Universal Robots URScript: FaiChun_9 Jan_3.script

def Machining1():
  # Default parameters:
  global speed_ms = 0.03
  global speed_rads = 0.75
  global accel_mss = 3
  global accel_radss = 1.2
  global blend_radius_m = 0.0003

  # Add subprograms here
  # Start of main program
  # Program generated by RoboDK v5.6.8 for UR10e on 09/01/2025 16:15:55
  # Using nominal kinematics.
  blend_radius_m = 0.0003
  speed_ms = 0.03
  # set_reference(p[0.335000, -0.060000, 0.000000, 0.000000, 0.000000, 0.000000])
  set_tcp(p[0.000000, 0.000000, 0.252000, 0.000000, 0.000000, 0.000000])
  # Show Tool
  movej([0.602689, -1.119966, -2.613047, -0.979376, 1.570796, 2.173486],accel_radss,speed_rads,0,blend_radius_m)
  movel([0.602689, -1.179994, -2.651340, -0.881054, 1.570796, 2.173486],accel_mss,speed_ms,0,blend_radius_m)
  #SetTool1
  #M_RunCode6
  #SetRPM60000
  speed_ms = 0.03
  #M_RunCode3
  movel([0.602689, -1.207513, -2.665873, -0.839003, 1.570796, 2.173486],accel_mss,speed_ms,0,blend_radius_m)
  speed_ms = 0.003
  movel([0.602689, -1.214750, -2.669441, -0.828198, 1.570796, 2.173486],accel_mss,speed_ms,0,blend_radius_m)
  speed_ms = 0.007
  movel([0.623056, -1.305978, -2.619553, -0.786857, 1.570796, 2.193852],accel_mss,speed_ms,0,blend_radius_m)
  movel([0.614868, -1.310439, -2.616847, -0.785103, 1.570796, 2.185664],accel_mss,speed_ms,0,blend_radius_m)
  movel([0.615927, -1.315223, -2.613916, -0.783250, 1.570796, 2.186723],accel_mss,speed_ms,0,blend_radius_m)
  movel([0.618034, -1.314081, -2.614619, -0.783689, 1.570796, 2.188830],accel_mss,speed_ms,0,blend_radius_m)
  movel([0.617346, -1.310924, -2.616551, -0.784913, 1.570796, 2.188143],accel_mss,speed_ms,0,blend_radius_m)
  movel([0.623401, -1.307643, -2.618547, -0.786200, 1.570796, 2.194198],accel_mss,speed_ms,0,blend_radius_m)
  movel([0.623560, -1.308410, -2.618081, -0.785898, 1.570796, 2.194357],accel_mss,speed_ms,0,blend_radius_m)
  movel([0.624387, -1.312349, -2.615681, -0.784359, 1.570796, 2.195184],accel_mss,speed_ms,0,blend_radius_m)
  movel([0.620317, -1.314540, -2.614336, -0.783512, 1.570796, 2.191113],accel_mss,speed_ms,0,blend_radius_m)
  movel([0.620668, -1.316175, -2.613329, -0.782885, 1.570796, 2.191464],accel_mss,speed_ms,0,blend_radius_m)
  movel([0.624731, -1.313996, -2.614671, -0.783722, 1.570796, 2.195527],accel_mss,speed_ms,0,blend_radius_m)
  movel([0.625701, -1.318667, -2.611788, -0.781935, 1.570796, 2.196498],accel_mss,speed_ms,0,blend_radius_m)
  movel([0.621661, -1.320822, -2.610447, -0.781120, 1.570796, 2.192457],accel_mss,speed_ms,0,blend_radius_m)
  movel([0.622322, -1.323943, -2.608496, -0.779950, 1.570796, 2.193118],accel_mss,speed_ms,0,blend_radius_m)
  movel([0.616386, -1.327108, -2.606503, -0.778778, 1.570796, 2.187182],accel_mss,speed_ms,0,blend_radius_m)
  movel([0.615701, -1.324013, -2.608452, -0.779924, 1.570796, 2.186497],accel_mss,speed_ms,0,blend_radius_m)
  movel([0.613619, -1.325132, -2.607748, -0.779508, 1.570796, 2.184416],accel_mss,speed_ms,0,blend_radius_m)
  movel([0.614310, -1.328222, -2.605799, -0.778369, 1.570796, 2.185106],accel_mss,speed_ms,0,blend_radius_m)
  movel([0.609368, -1.330876, -2.604114, -0.777400, 1.570796, 2.180164],accel_mss,speed_ms,0,blend_radius_m)
  movel([0.608412, -1.331392, -2.603784, -0.777212, 1.570796, 2.179209],accel_mss,speed_ms,0,blend_radius_m)
  movel([0.607352, -1.326855, -2.606663, -0.778871, 1.570796, 2.178148],accel_mss,speed_ms,0,blend_radius_m)
  movel([0.611354, -1.324685, -2.608029, -0.779674, 1.570796, 2.182150],accel_mss,speed_ms,0,blend_radius_m)
  movel([0.610987, -1.323080, -2.609036, -0.780272, 1.570796, 2.181784],accel_mss,speed_ms,0,blend_radius_m)
  movel([0.604903, -1.326389, -2.606957, -0.779043, 1.570796, 2.175699],accel_mss,speed_ms,0,blend_radius_m)
  movel([0.606349, -1.332504, -2.603075, -0.776810, 1.570796, 2.177146],accel_mss,speed_ms,0,blend_radius_m)
  movel([0.503740, -1.390840, -2.563439, -0.758110, 1.570796, 2.074536],accel_mss,speed_ms,0,blend_radius_m)
  movel([0.410742, -1.448915, -2.519079, -0.744396, 1.570796, 1.981539],accel_mss,speed_ms,0,blend_radius_m)
  movel([0.408155, -1.444408, -2.522703, -0.745278, 1.570796, 1.978951],accel_mss,speed_ms,0,blend_radius_m)
  movel([0.403196, -1.447676, -2.520078, -0.744635, 1.570796, 1.973993],accel_mss,speed_ms,0,blend_radius_m)
  movel([0.403874, -1.448837, -2.519141, -0.744410, 1.570796, 1.974671],accel_mss,speed_ms,0,blend_radius_m)
  movel([0.407131, -1.446693, -2.520869, -0.744827, 1.570796, 1.977928],accel_mss,speed_ms,0,blend_radius_m)
  movel([0.409046, -1.450019, -2.518186, -0.744184, 1.570796, 1.979842],accel_mss,speed_ms,0,blend_radius_m)
  movel([0.408262, -1.450531, -2.517771, -0.744086, 1.570796, 1.979059],accel_mss,speed_ms,0,blend_radius_m)
  movel([0.404240, -1.453169, -2.515629, -0.743591, 1.570796, 1.975036],accel_mss,speed_ms,0,blend_radius_m)
  movel([0.402940, -1.450940, -2.517440, -0.744009, 1.570796, 1.973737],accel_mss,speed_ms,0,blend_radius_m)
  movel([0.401260, -1.452049, -2.516540, -0.743800, 1.570796, 1.972056],accel_mss,speed_ms,0,blend_radius_m)
  movel([0.402562, -1.454272, -2.514730, -0.743387, 1.570796, 1.973359],accel_mss,speed_ms,0,blend_radius_m)
  movel([0.397796, -1.457416, -2.512158, -0.742815, 1.570796, 1.968593],accel_mss,speed_ms,0,blend_radius_m)
  movel([0.396480, -1.455213, -2.513962, -0.743214, 1.570796, 1.967277],accel_mss,speed_ms,0,blend_radius_m)
  movel([0.393271, -1.457346, -2.512215, -0.742828, 1.570796, 1.964067],accel_mss,speed_ms,0,blend_radius_m)
  movel([0.391300, -1.454096, -2.514874, -0.743419, 1.570796, 1.962097],accel_mss,speed_ms,0,blend_radius_m)
  movel([0.394521, -1.451944, -2.516626, -0.743820, 1.570796, 1.965317],accel_mss,speed_ms,0,blend_radius_m)
  movel([0.393830, -1.450797, -2.517556, -0.744036, 1.570796, 1.964626],accel_mss,speed_ms,0,blend_radius_m)
  movel([0.390606, -1.452954, -2.515804, -0.743631, 1.570796, 1.961403],accel_mss,speed_ms,0,blend_radius_m)
  movel([0.388934, -1.450227, -2.518017, -0.744144, 1.570796, 1.959730],accel_mss,speed_ms,0,blend_radius_m)
  movel([0.388611, -1.449697, -2.518446, -0.744245, 1.570796, 1.959407],accel_mss,speed_ms,0,blend_radius_m)
  movel([0.393406, -1.446476, -2.521044, -0.744869, 1.570796, 1.964202],accel_mss,speed_ms,0,blend_radius_m)
  movel([0.394744, -1.448694, -2.519257, -0.744438, 1.570796, 1.965540],accel_mss,speed_ms,0,blend_radius_m)
  movel([0.396427, -1.447570, -2.520164, -0.744656, 1.570796, 1.967224],accel_mss,speed_ms,0,blend_radius_m)
  movel([0.394398, -1.444188, -2.522879, -0.745322, 1.570796, 1.965194],accel_mss,speed_ms,0,blend_radius_m)
  movel([0.387908, -1.448555, -2.519369, -0.744465, 1.570796, 1.958704],accel_mss,speed_ms,0,blend_radius_m)
  movel([0.387580, -1.448026, -2.519796, -0.744567, 1.570796, 1.958376],accel_mss,speed_ms,0,blend_radius_m)
  movel([0.348021, -1.388149, -2.565374, -0.758866, 1.570796, 1.918817],accel_mss,speed_ms,0,blend_radius_m)
  movel([0.300929, -1.326689, -2.606767, -0.778932, 1.570796, 1.871725],accel_mss,speed_ms,0,blend_radius_m)
  movel([0.308156, -1.320668, -2.610543, -0.781178, 1.570796, 1.878952],accel_mss,speed_ms,0,blend_radius_m)
  movel([0.305290, -1.317157, -2.612722, -0.782509, 1.570796, 1.876086],accel_mss,speed_ms,0,blend_radius_m)
  movel([0.303402, -1.318735, -2.611745, -0.781909, 1.570796, 1.874198],accel_mss,speed_ms,0,blend_radius_m)
  movel([0.305295, -1.321037, -2.610313, -0.781039, 1.570796, 1.876092],accel_mss,speed_ms,0,blend_radius_m)
  movel([0.299947, -1.325499, -2.607518, -0.779372, 1.570796, 1.870743],accel_mss,speed_ms,0,blend_radius_m)
  movel([0.299492, -1.324951, -2.607863, -0.779576, 1.570796, 1.870288],accel_mss,speed_ms,0,blend_radius_m)
  movel([0.297126, -1.322128, -2.609632, -0.780629, 1.570796, 1.867922],accel_mss,speed_ms,0,blend_radius_m)
  movel([0.300740, -1.319092, -2.611523, -0.781773, 1.570796, 1.871536],accel_mss,speed_ms,0,blend_radius_m)
  movel([0.299747, -1.317902, -2.612261, -0.782225, 1.570796, 1.870544],accel_mss,speed_ms,0,blend_radius_m)
  movel([0.296130, -1.320947, -2.610369, -0.781072, 1.570796, 1.866927],accel_mss,speed_ms,0,blend_radius_m)
  movel([0.293273, -1.317580, -2.612461, -0.782348, 1.570796, 1.864069],accel_mss,speed_ms,0,blend_radius_m)
  movel([0.296899, -1.314508, -2.614356, -0.783525, 1.570796, 1.867695],accel_mss,speed_ms,0,blend_radius_m)
  movel([0.294961, -1.312214, -2.615763, -0.784412, 1.570796, 1.865757],accel_mss,speed_ms,0,blend_radius_m)
  movel([0.300378, -1.307616, -2.618562, -0.786210, 1.570796, 1.871174],accel_mss,speed_ms,0,blend_radius_m)
  movel([0.302307, -1.309936, -2.617154, -0.785299, 1.570796, 1.873103],accel_mss,speed_ms,0,blend_radius_m)
  movel([0.304213, -1.308328, -2.618131, -0.785930, 1.570796, 1.875010],accel_mss,speed_ms,0,blend_radius_m)
  movel([0.302287, -1.305999, -2.619541, -0.786849, 1.570796, 1.873084],accel_mss,speed_ms,0,blend_radius_m)
  movel([0.306872, -1.302122, -2.621872, -0.788396, 1.570796, 1.877668],accel_mss,speed_ms,0,blend_radius_m)
  movel([0.307765, -1.301370, -2.622322, -0.788698, 1.570796, 1.878562],accel_mss,speed_ms,0,blend_radius_m)
  movel([0.310601, -1.304861, -2.620227, -0.787301, 1.570796, 1.881398],accel_mss,speed_ms,0,blend_radius_m)
  movel([0.306907, -1.307961, -2.618354, -0.786074, 1.570796, 1.877703],accel_mss,speed_ms,0,blend_radius_m)
  movel([0.307897, -1.309175, -2.617616, -0.785597, 1.570796, 1.878694],accel_mss,speed_ms,0,blend_radius_m)
  movel([0.313513, -1.304476, -2.620459, -0.787454, 1.570796, 1.884309],accel_mss,speed_ms,0,blend_radius_m)
  movel([0.309700, -1.299738, -2.623295, -0.789356, 1.570796, 1.880496],accel_mss,speed_ms,0,blend_radius_m)
  movel([0.418732, -1.210473, -2.671537, -0.830378, 1.570796, 1.989529],accel_mss,speed_ms,0,blend_radius_m)
  movel([0.544562, -1.113334, -2.713941, -0.885114, 1.570796, 2.115358],accel_mss,speed_ms,0,blend_radius_m)
  movel([0.545777, -1.112427, -2.714293, -0.885669, 1.570796, 2.116573],accel_mss,speed_ms,0,blend_radius_m)
  movel([0.548232, -1.120070, -2.711305, -0.881014, 1.570796, 2.119029],accel_mss,speed_ms,0,blend_radius_m)
  movel([0.555880, -1.114419, -2.713519, -0.884450, 1.570796, 2.126677],accel_mss,speed_ms,0,blend_radius_m)
  movel([0.555266, -1.112413, -2.714298, -0.885678, 1.570796, 2.126062],accel_mss,speed_ms,0,blend_radius_m)
  movel([0.550215, -1.116152, -2.712844, -0.883393, 1.570796, 2.121011],accel_mss,speed_ms,0,blend_radius_m)
  movel([0.548415, -1.110463, -2.715052, -0.886874, 1.570796, 2.119211],accel_mss,speed_ms,0,blend_radius_m)
  movel([0.549632, -1.109554, -2.715402, -0.887433, 1.570796, 2.120428],accel_mss,speed_ms,0,blend_radius_m)
  movel([0.555951, -1.104840, -2.717204, -0.890344, 1.570796, 2.126748],accel_mss,speed_ms,0,blend_radius_m)
  movel([0.557137, -1.108742, -2.715714, -0.887933, 1.570796, 2.127934],accel_mss,speed_ms,0,blend_radius_m)
  movel([0.559782, -1.106785, -2.716463, -0.889141, 1.570796, 2.130578],accel_mss,speed_ms,0,blend_radius_m)
  movel([0.558607, -1.102864, -2.717954, -0.891571, 1.570796, 2.129404],accel_mss,speed_ms,0,blend_radius_m)
  movel([0.566225, -1.097212, -2.720078, -0.895099, 1.570796, 2.137021],accel_mss,speed_ms,0,blend_radius_m)
  movel([0.567373, -1.101184, -2.718589, -0.892617, 1.570796, 2.138169],accel_mss,speed_ms,0,blend_radius_m)
  movel([0.572529, -1.097390, -2.720012, -0.894987, 1.570796, 2.143326],accel_mss,speed_ms,0,blend_radius_m)
  movel([0.574176, -1.103301, -2.717789, -0.891299, 1.570796, 2.144972],accel_mss,speed_ms,0,blend_radius_m)
  movel([0.569046, -1.107043, -2.716364, -0.888981, 1.570796, 2.139842],accel_mss,speed_ms,0,blend_radius_m)
  movel([0.569628, -1.109089, -2.715581, -0.887720, 1.570796, 2.140424],accel_mss,speed_ms,0,blend_radius_m)
  movel([0.574746, -1.105365, -2.717005, -0.890019, 1.570796, 2.145542],accel_mss,speed_ms,0,blend_radius_m)
  movel([0.576356, -1.111236, -2.714753, -0.886399, 1.570796, 2.147153],accel_mss,speed_ms,0,blend_radius_m)
  movel([0.568840, -1.116662, -2.712644, -0.883082, 1.570796, 2.139637],accel_mss,speed_ms,0,blend_radius_m)
  movel([0.567720, -1.112757, -2.714165, -0.885467, 1.570796, 2.138516],accel_mss,speed_ms,0,blend_radius_m)
  movel([0.565088, -1.114673, -2.713421, -0.884296, 1.570796, 2.135884],accel_mss,speed_ms,0,blend_radius_m)
  movel([0.566799, -1.120576, -2.711106, -0.880707, 1.570796, 2.137595],accel_mss,speed_ms,0,blend_radius_m)
  movel([0.576916, -1.113286, -2.713960, -0.885143, 1.570796, 2.147712],accel_mss,speed_ms,0,blend_radius_m)
  movel([0.602689, -1.214750, -2.669441, -0.828198, 1.570796, 2.173486],accel_mss,speed_ms,0,blend_radius_m)
  speed_ms = 0.003
  movel([0.602689, -1.207513, -2.665873, -0.839003, 1.570796, 2.173486],accel_mss,speed_ms,0,blend_radius_m)
  speed_ms = 0.03
  movel([0.602689, -1.179994, -2.651340, -0.881054, 1.570796, 2.173486],accel_mss,speed_ms,0,blend_radius_m)
  #M_RunCode9
  movel([0.550774, -1.125627, -2.675411, -0.911351, 1.570796, 2.121570],accel_mss,speed_ms,0,blend_radius_m)
  #M_RunCode3
  movel([0.550774, -1.153488, -2.690658, -0.868243, 1.570796, 2.121570],accel_mss,speed_ms,0,blend_radius_m)
  speed_ms = 0.003
  movel([0.550774, -1.160850, -2.694409, -0.857131, 1.570796, 2.121570],accel_mss,speed_ms,0,blend_radius_m)
  speed_ms = 0.007
  movel([0.548561, -1.162804, -2.693557, -0.856028, 1.570796, 2.119358],accel_mss,speed_ms,0,blend_radius_m)
  movel([0.546305, -1.164169, -2.692960, -0.855260, 1.570796, 2.117101],accel_mss,speed_ms,0,blend_radius_m)
  movel([0.543998, -1.164956, -2.692615, -0.854818, 1.570796, 2.114794],accel_mss,speed_ms,0,blend_radius_m)
  movel([0.541636, -1.165162, -2.692525, -0.854702, 1.570796, 2.112432],accel_mss,speed_ms,0,blend_radius_m)
  movel([0.539730, -1.164842, -2.692665, -0.854882, 1.570796, 2.110526],accel_mss,speed_ms,0,blend_radius_m)
  movel([0.538223, -1.164013, -2.693029, -0.855348, 1.570796, 2.109019],accel_mss,speed_ms,0,blend_radius_m)
  movel([0.537059, -1.162815, -2.693552, -0.856021, 1.570796, 2.107855],accel_mss,speed_ms,0,blend_radius_m)
  movel([0.536184, -1.161380, -2.694178, -0.856831, 1.570796, 2.106980],accel_mss,speed_ms,0,blend_radius_m)
  movel([0.534689, -1.157276, -2.695956, -0.859157, 1.570796, 2.105485],accel_mss,speed_ms,0,blend_radius_m)
  movel([0.533234, -1.153410, -2.697615, -0.861364, 1.570796, 2.104030],accel_mss,speed_ms,0,blend_radius_m)
  movel([0.532433, -1.152087, -2.698179, -0.862123, 1.570796, 2.103229],accel_mss,speed_ms,0,blend_radius_m)
  movel([0.531381, -1.150992, -2.698644, -0.862753, 1.570796, 2.102177],accel_mss,speed_ms,0,blend_radius_m)
  movel([0.530038, -1.150250, -2.698959, -0.863179, 1.570796, 2.100835],accel_mss,speed_ms,0,blend_radius_m)
  movel([0.528363, -1.149991, -2.699069, -0.863329, 1.570796, 2.099159],accel_mss,speed_ms,0,blend_radius_m)
  movel([0.527809, -1.151106, -2.698596, -0.862687, 1.570796, 2.098605],accel_mss,speed_ms,0,blend_radius_m)
  movel([0.526408, -1.154185, -2.697283, -0.860921, 1.570796, 2.097204],accel_mss,speed_ms,0,blend_radius_m)
  movel([0.525462, -1.156876, -2.696128, -0.859385, 1.570796, 2.096259],accel_mss,speed_ms,0,blend_radius_m)
  movel([0.524967, -1.159182, -2.695132, -0.858075, 1.570796, 2.095763],accel_mss,speed_ms,0,blend_radius_m)
  movel([0.524917, -1.161112, -2.694295, -0.856982, 1.570796, 2.095713],accel_mss,speed_ms,0,blend_radius_m)
  movel([0.525250, -1.162687, -2.693608, -0.856093, 1.570796, 2.096047],accel_mss,speed_ms,0,blend_radius_m)
  movel([0.525915, -1.163932, -2.693064, -0.855393, 1.570796, 2.096711],accel_mss,speed_ms,0,blend_radius_m)
  movel([0.526910, -1.164844, -2.692664, -0.854881, 1.570796, 2.097706],accel_mss,speed_ms,0,blend_radius_m)
  movel([0.528231, -1.165431, -2.692406, -0.854551, 1.570796, 2.099027],accel_mss,speed_ms,0,blend_radius_m)
  movel([0.519926, -1.165324, -2.692454, -0.854612, 1.570796, 2.090722],accel_mss,speed_ms,0,blend_radius_m)
  movel([0.534681, -1.135580, -2.705071, -0.871737, 1.570796, 2.105477],accel_mss,speed_ms,0,blend_radius_m)
  movel([0.535536, -1.135588, -2.705068, -0.871733, 1.570796, 2.106332],accel_mss,speed_ms,0,blend_radius_m)
  movel([0.537525, -1.135957, -2.704917, -0.871515, 1.570796, 2.108321],accel_mss,speed_ms,0,blend_radius_m)
  movel([0.539121, -1.137030, -2.704477, -0.870882, 1.570796, 2.109917],accel_mss,speed_ms,0,blend_radius_m)
  movel([0.540368, -1.138595, -2.703833, -0.869961, 1.570796, 2.111164],accel_mss,speed_ms,0,blend_radius_m)
  movel([0.541307, -1.140440, -2.703070, -0.868879, 1.570796, 2.112103],accel_mss,speed_ms,0,blend_radius_m)
  movel([0.543134, -1.145919, -2.700786, -0.865684, 1.570796, 2.113931],accel_mss,speed_ms,0,blend_radius_m)
  movel([0.544743, -1.151028, -2.698629, -0.862732, 1.570796, 2.115539],accel_mss,speed_ms,0,blend_radius_m)
  movel([0.545581, -1.152750, -2.697896, -0.861743, 1.570796, 2.116377],accel_mss,speed_ms,0,blend_radius_m)
  movel([0.546665, -1.154185, -2.697283, -0.860921, 1.570796, 2.117461],accel_mss,speed_ms,0,blend_radius_m)
  movel([0.548025, -1.155169, -2.696862, -0.860358, 1.570796, 2.118821],accel_mss,speed_ms,0,blend_radius_m)
  movel([0.549683, -1.155544, -2.696701, -0.860144, 1.570796, 2.120479],accel_mss,speed_ms,0,blend_radius_m)
  movel([0.552028, -1.155227, -2.696837, -0.860325, 1.570796, 2.122824],accel_mss,speed_ms,0,blend_radius_m)
  movel([0.553135, -1.154766, -2.697035, -0.860589, 1.570796, 2.123932],accel_mss,speed_ms,0,blend_radius_m)
  movel([0.554203, -1.154097, -2.697321, -0.860971, 1.570796, 2.125000],accel_mss,speed_ms,0,blend_radius_m)
  movel([0.556059, -1.152398, -2.698046, -0.861944, 1.570796, 2.126856],accel_mss,speed_ms,0,blend_radius_m)
  movel([0.557429, -1.150391, -2.698899, -0.863098, 1.570796, 2.128225],accel_mss,speed_ms,0,blend_radius_m)
  movel([0.558020, -1.149017, -2.699481, -0.863891, 1.570796, 2.128816],accel_mss,speed_ms,0,blend_radius_m)
  movel([0.558180, -1.147987, -2.699916, -0.864486, 1.570796, 2.128976],accel_mss,speed_ms,0,blend_radius_m)
  movel([0.557957, -1.147333, -2.700192, -0.864864, 1.570796, 2.128753],accel_mss,speed_ms,0,blend_radius_m)
  movel([0.557399, -1.147097, -2.700291, -0.865001, 1.570796, 2.128195],accel_mss,speed_ms,0,blend_radius_m)
  movel([0.556151, -1.147552, -2.700100, -0.864738, 1.570796, 2.126947],accel_mss,speed_ms,0,blend_radius_m)
  movel([0.554911, -1.148103, -2.699867, -0.864419, 1.570796, 2.125708],accel_mss,speed_ms,0,blend_radius_m)
  movel([0.553550, -1.148272, -2.699796, -0.864321, 1.570796, 2.124347],accel_mss,speed_ms,0,blend_radius_m)
  movel([0.552254, -1.147868, -2.699966, -0.864555, 1.570796, 2.123050],accel_mss,speed_ms,0,blend_radius_m)
  movel([0.551694, -1.146779, -2.700425, -0.865185, 1.570796, 2.122490],accel_mss,speed_ms,0,blend_radius_m)
  movel([0.551802, -1.145219, -2.701079, -0.866090, 1.570796, 2.122598],accel_mss,speed_ms,0,blend_radius_m)
  movel([0.552503, -1.143409, -2.701836, -0.867144, 1.570796, 2.123299],accel_mss,speed_ms,0,blend_radius_m)
  movel([0.553665, -1.141608, -2.702586, -0.868195, 1.570796, 2.124461],accel_mss,speed_ms,0,blend_radius_m)
  movel([0.555150, -1.140087, -2.703216, -0.869085, 1.570796, 2.125946],accel_mss,speed_ms,0,blend_radius_m)
  movel([0.556809, -1.139065, -2.703639, -0.869685, 1.570796, 2.127606],accel_mss,speed_ms,0,blend_radius_m)
  movel([0.558480, -1.138768, -2.703761, -0.869860, 1.570796, 2.129276],accel_mss,speed_ms,0,blend_radius_m)
  movel([0.559682, -1.139024, -2.703656, -0.869709, 1.570796, 2.130479],accel_mss,speed_ms,0,blend_radius_m)
  movel([0.560510, -1.139683, -2.703383, -0.869322, 1.570796, 2.131306],accel_mss,speed_ms,0,blend_radius_m)
  movel([0.560959, -1.140749, -2.702942, -0.868698, 1.570796, 2.131755],accel_mss,speed_ms,0,blend_radius_m)
  movel([0.561036, -1.142210, -2.702335, -0.867843, 1.570796, 2.131832],accel_mss,speed_ms,0,blend_radius_m)
  movel([0.560782, -1.143971, -2.701602, -0.866816, 1.570796, 2.131579],accel_mss,speed_ms,0,blend_radius_m)
  movel([0.560231, -1.145930, -2.700781, -0.865677, 1.570796, 2.131028],accel_mss,speed_ms,0,blend_radius_m)
  movel([0.558257, -1.150429, -2.698884, -0.863077, 1.570796, 2.129054],accel_mss,speed_ms,0,blend_radius_m)
  movel([0.556625, -1.153304, -2.697660, -0.861425, 1.570796, 2.127421],accel_mss,speed_ms,0,blend_radius_m)
  movel([0.554835, -1.155999, -2.696505, -0.859885, 1.570796, 2.125631],accel_mss,speed_ms,0,blend_radius_m)
  movel([0.552885, -1.158510, -2.695423, -0.858456, 1.570796, 2.123681],accel_mss,speed_ms,0,blend_radius_m)
  movel([0.550774, -1.160850, -2.694409, -0.857131, 1.570796, 2.121570],accel_mss,speed_ms,0,blend_radius_m)
  speed_ms = 0.003
  movel([0.550774, -1.153488, -2.690658, -0.868243, 1.570796, 2.121570],accel_mss,speed_ms,0,blend_radius_m)
  speed_ms = 0.03
  movel([0.550774, -1.125627, -2.675411, -0.911351, 1.570796, 2.121570],accel_mss,speed_ms,0,blend_radius_m)
  #M_RunCode9
  movel([0.538556, -1.144823, -2.667250, -0.900316, 1.570796, 2.109352],accel_mss,speed_ms,0,blend_radius_m)
  #M_RunCode3
  movel([0.538556, -1.172591, -2.682246, -0.857552, 1.570796, 2.109352],accel_mss,speed_ms,0,blend_radius_m)
  speed_ms = 0.003
  movel([0.538556, -1.179915, -2.685933, -0.846541, 1.570796, 2.109352],accel_mss,speed_ms,0,blend_radius_m)
  speed_ms = 0.007
  movel([0.539812, -1.180524, -2.685656, -0.846209, 1.570796, 2.110609],accel_mss,speed_ms,0,blend_radius_m)
  movel([0.540517, -1.181326, -2.685290, -0.845773, 1.570796, 2.111313],accel_mss,speed_ms,0,blend_radius_m)
  movel([0.540674, -1.182325, -2.684834, -0.845230, 1.570796, 2.111471],accel_mss,speed_ms,0,blend_radius_m)
  movel([0.540282, -1.183515, -2.684289, -0.844585, 1.570796, 2.111078],accel_mss,speed_ms,0,blend_radius_m)
  movel([0.539454, -1.184688, -2.683751, -0.843950, 1.570796, 2.110251],accel_mss,speed_ms,0,blend_radius_m)
  movel([0.538299, -1.185627, -2.683319, -0.843443, 1.570796, 2.109096],accel_mss,speed_ms,0,blend_radius_m)
  movel([0.536822, -1.186334, -2.682993, -0.843062, 1.570796, 2.107618],accel_mss,speed_ms,0,blend_radius_m)
  movel([0.535012, -1.186818, -2.682769, -0.842802, 1.570796, 2.105809],accel_mss,speed_ms,0,blend_radius_m)
  movel([0.530250, -1.187319, -2.682538, -0.842532, 1.570796, 2.101046],accel_mss,speed_ms,0,blend_radius_m)
  movel([0.523846, -1.187356, -2.682521, -0.842512, 1.570796, 2.094643],accel_mss,speed_ms,0,blend_radius_m)
  movel([0.517633, -1.187006, -2.682682, -0.842700, 1.570796, 2.088430],accel_mss,speed_ms,0,blend_radius_m)
  movel([0.513485, -1.186284, -2.683016, -0.843089, 1.570796, 2.084281],accel_mss,speed_ms,0,blend_radius_m)
  movel([0.512201, -1.185722, -2.683275, -0.843392, 1.570796, 2.082997],accel_mss,speed_ms,0,blend_radius_m)
  movel([0.511463, -1.184959, -2.683626, -0.843803, 1.570796, 2.082259],accel_mss,speed_ms,0,blend_radius_m)
  movel([0.511270, -1.183986, -2.684073, -0.844330, 1.570796, 2.082067],accel_mss,speed_ms,0,blend_radius_m)
  movel([0.511631, -1.182800, -2.684617, -0.844972, 1.570796, 2.082427],accel_mss,speed_ms,0,blend_radius_m)
  movel([0.512434, -1.181618, -2.685157, -0.845614, 1.570796, 2.083230],accel_mss,speed_ms,0,blend_radius_m)
  movel([0.513582, -1.180651, -2.685598, -0.846140, 1.570796, 2.084378],accel_mss,speed_ms,0,blend_radius_m)
  movel([0.515069, -1.179904, -2.685938, -0.846547, 1.570796, 2.085865],accel_mss,speed_ms,0,blend_radius_m)
  movel([0.516901, -1.179372, -2.686179, -0.846838, 1.570796, 2.087698],accel_mss,speed_ms,0,blend_radius_m)
  movel([0.521734, -1.178775, -2.686450, -0.847164, 1.570796, 2.092531],accel_mss,speed_ms,0,blend_radius_m)
  movel([0.528212, -1.178691, -2.686488, -0.847210, 1.570796, 2.099008],accel_mss,speed_ms,0,blend_radius_m)
  movel([0.534440, -1.179094, -2.686306, -0.846989, 1.570796, 2.105236],accel_mss,speed_ms,0,blend_radius_m)
  movel([0.538556, -1.179915, -2.685933, -0.846541, 1.570796, 2.109352],accel_mss,speed_ms,0,blend_radius_m)
  speed_ms = 0.003
  movel([0.538556, -1.172591, -2.682246, -0.857552, 1.570796, 2.109352],accel_mss,speed_ms,0,blend_radius_m)
  speed_ms = 0.03
  movel([0.538556, -1.144823, -2.667250, -0.900316, 1.570796, 2.109352],accel_mss,speed_ms,0,blend_radius_m)
  #M_RunCode9
  movel([0.542858, -1.143015, -2.668034, -0.901339, 1.570796, 2.113654],accel_mss,speed_ms,0,blend_radius_m)
  #M_RunCode3
  movel([0.542858, -1.170793, -2.683054, -0.858542, 1.570796, 2.113654],accel_mss,speed_ms,0,blend_radius_m)
  speed_ms = 0.003
  movel([0.542858, -1.178121, -2.686746, -0.847521, 1.570796, 2.113654],accel_mss,speed_ms,0,blend_radius_m)
  speed_ms = 0.007
  movel([0.542513, -1.179848, -2.685963, -0.846578, 1.570796, 2.113310],accel_mss,speed_ms,0,blend_radius_m)
  movel([0.541905, -1.181659, -2.685138, -0.845592, 1.570796, 2.112701],accel_mss,speed_ms,0,blend_radius_m)
  movel([0.541037, -1.183547, -2.684275, -0.844567, 1.570796, 2.111833],accel_mss,speed_ms,0,blend_radius_m)
  movel([0.539959, -1.185423, -2.683413, -0.843553, 1.570796, 2.110755],accel_mss,speed_ms,0,blend_radius_m)
  movel([0.538720, -1.187190, -2.682598, -0.842602, 1.570796, 2.109516],accel_mss,speed_ms,0,blend_radius_m)
  movel([0.537321, -1.188846, -2.681830, -0.841713, 1.570796, 2.108117],accel_mss,speed_ms,0,blend_radius_m)
  movel([0.535761, -1.190396, -2.681110, -0.840884, 1.570796, 2.106557],accel_mss,speed_ms,0,blend_radius_m)
  movel([0.534059, -1.191809, -2.680450, -0.840129, 1.570796, 2.104855],accel_mss,speed_ms,0,blend_radius_m)
  movel([0.532235, -1.193051, -2.679869, -0.839469, 1.570796, 2.103031],accel_mss,speed_ms,0,blend_radius_m)
  movel([0.530283, -1.194130, -2.679363, -0.838896, 1.570796, 2.101080],accel_mss,speed_ms,0,blend_radius_m)
  movel([0.528204, -1.195044, -2.678933, -0.838412, 1.570796, 2.099000],accel_mss,speed_ms,0,blend_radius_m)
  movel([0.526038, -1.195762, -2.678595, -0.838032, 1.570796, 2.096834],accel_mss,speed_ms,0,blend_radius_m)
  movel([0.523816, -1.196259, -2.678360, -0.837770, 1.570796, 2.094612],accel_mss,speed_ms,0,blend_radius_m)
  movel([0.521541, -1.196533, -2.678231, -0.837625, 1.570796, 2.092337],accel_mss,speed_ms,0,blend_radius_m)
  movel([0.519210, -1.196586, -2.678206, -0.837598, 1.570796, 2.090007],accel_mss,speed_ms,0,blend_radius_m)
  movel([0.516986, -1.196422, -2.678283, -0.837684, 1.570796, 2.087782],accel_mss,speed_ms,0,blend_radius_m)
  movel([0.515037, -1.196045, -2.678461, -0.837883, 1.570796, 2.085833],accel_mss,speed_ms,0,blend_radius_m)
  movel([0.513361, -1.195453, -2.678741, -0.838196, 1.570796, 2.084157],accel_mss,speed_ms,0,blend_radius_m)
  movel([0.511958, -1.194647, -2.679120, -0.838622, 1.570796, 2.082755],accel_mss,speed_ms,0,blend_radius_m)
  movel([0.510836, -1.193654, -2.679587, -0.839149, 1.570796, 2.081632],accel_mss,speed_ms,0,blend_radius_m)
  movel([0.509996, -1.192506, -2.680125, -0.839759, 1.570796, 2.080792],accel_mss,speed_ms,0,blend_radius_m)
  movel([0.509441, -1.191204, -2.680733, -0.840452, 1.570796, 2.080237],accel_mss,speed_ms,0,blend_radius_m)
  movel([0.509173, -1.189740, -2.681415, -0.841234, 1.570796, 2.079969],accel_mss,speed_ms,0,blend_radius_m)
  movel([0.509180, -1.188151, -2.682153, -0.842086, 1.570796, 2.079976],accel_mss,speed_ms,0,blend_radius_m)
  movel([0.509453, -1.186465, -2.682933, -0.842992, 1.570796, 2.080250],accel_mss,speed_ms,0,blend_radius_m)
  movel([0.509999, -1.184678, -2.683755, -0.843955, 1.570796, 2.080796],accel_mss,speed_ms,0,blend_radius_m)
  movel([0.510812, -1.182794, -2.684620, -0.844976, 1.570796, 2.081609],accel_mss,speed_ms,0,blend_radius_m)
  movel([0.511849, -1.180908, -2.685481, -0.846000, 1.570796, 2.082645],accel_mss,speed_ms,0,blend_radius_m)
  movel([0.513063, -1.179109, -2.686299, -0.846981, 1.570796, 2.083859],accel_mss,speed_ms,0,blend_radius_m)
  movel([0.514458, -1.177407, -2.687070, -0.847913, 1.570796, 2.085254],accel_mss,speed_ms,0,blend_radius_m)
  movel([0.516032, -1.175798, -2.687795, -0.848796, 1.570796, 2.086828],accel_mss,speed_ms,0,blend_radius_m)
  movel([0.517764, -1.174315, -2.688462, -0.849612, 1.570796, 2.088560],accel_mss,speed_ms,0,blend_radius_m)
  movel([0.519630, -1.172997, -2.689052, -0.850340, 1.570796, 2.090427],accel_mss,speed_ms,0,blend_radius_m)
  movel([0.521632, -1.171848, -2.689565, -0.850976, 1.570796, 2.092428],accel_mss,speed_ms,0,blend_radius_m)
  movel([0.523768, -1.170863, -2.690004, -0.851522, 1.570796, 2.094564],accel_mss,speed_ms,0,blend_radius_m)
  movel([0.526000, -1.170084, -2.690351, -0.851954, 1.570796, 2.096797],accel_mss,speed_ms,0,blend_radius_m)
  movel([0.528286, -1.169540, -2.690592, -0.852257, 1.570796, 2.099082],accel_mss,speed_ms,0,blend_radius_m)
  movel([0.530626, -1.169238, -2.690726, -0.852425, 1.570796, 2.101422],accel_mss,speed_ms,0,blend_radius_m)
  movel([0.533019, -1.169178, -2.690753, -0.852458, 1.570796, 2.103815],accel_mss,speed_ms,0,blend_radius_m)
  movel([0.535288, -1.169357, -2.690673, -0.852359, 1.570796, 2.106084],accel_mss,speed_ms,0,blend_radius_m)
  movel([0.537266, -1.169770, -2.690490, -0.852129, 1.570796, 2.108062],accel_mss,speed_ms,0,blend_radius_m)
  movel([0.538952, -1.170414, -2.690204, -0.851771, 1.570796, 2.109748],accel_mss,speed_ms,0,blend_radius_m)
  movel([0.540346, -1.171286, -2.689816, -0.851287, 1.570796, 2.111143],accel_mss,speed_ms,0,blend_radius_m)
  movel([0.541445, -1.172352, -2.689341, -0.850697, 1.570796, 2.112241],accel_mss,speed_ms,0,blend_radius_m)
  movel([0.542243, -1.173571, -2.688795, -0.850023, 1.570796, 2.113039],accel_mss,speed_ms,0,blend_radius_m)
  movel([0.542738, -1.174948, -2.688178, -0.849264, 1.570796, 2.113535],accel_mss,speed_ms,0,blend_radius_m)
  movel([0.542938, -1.176477, -2.687489, -0.848423, 1.570796, 2.113734],accel_mss,speed_ms,0,blend_radius_m)
  movel([0.542858, -1.178121, -2.686746, -0.847521, 1.570796, 2.113654],accel_mss,speed_ms,0,blend_radius_m)
  speed_ms = 0.003
  movel([0.542858, -1.170793, -2.683054, -0.858542, 1.570796, 2.113654],accel_mss,speed_ms,0,blend_radius_m)
  speed_ms = 0.03
  movel([0.542858, -1.143015, -2.668034, -0.901339, 1.570796, 2.113654],accel_mss,speed_ms,0,blend_radius_m)
  #M_RunCode9
  movel([0.412645, -1.363842, -2.545198, -0.803350, 1.570796, 1.983441],accel_mss,speed_ms,0,blend_radius_m)
  #M_RunCode3
  movel([0.412645, -1.388740, -2.557323, -0.766326, 1.570796, 1.983441],accel_mss,speed_ms,0,blend_radius_m)
  speed_ms = 0.003
  movel([0.412645, -1.395201, -2.560281, -0.756906, 1.570796, 1.983441],accel_mss,speed_ms,0,blend_radius_m)
  speed_ms = 0.007
  movel([0.414245, -1.395440, -2.560107, -0.756841, 1.570796, 1.985042],accel_mss,speed_ms,0,blend_radius_m)
  movel([0.415609, -1.396135, -2.559602, -0.756652, 1.570796, 1.986405],accel_mss,speed_ms,0,blend_radius_m)
  movel([0.416748, -1.397147, -2.558864, -0.756378, 1.570796, 1.987545],accel_mss,speed_ms,0,blend_radius_m)
  movel([0.417677, -1.398344, -2.557989, -0.756056, 1.570796, 1.988473],accel_mss,speed_ms,0,blend_radius_m)
  movel([0.419680, -1.401911, -2.555369, -0.755109, 1.570796, 1.990477],accel_mss,speed_ms,0,blend_radius_m)
  movel([0.421479, -1.405241, -2.552907, -0.754241, 1.570796, 1.992276],accel_mss,speed_ms,0,blend_radius_m)
  movel([0.422316, -1.406367, -2.552070, -0.753952, 1.570796, 1.993112],accel_mss,speed_ms,0,blend_radius_m)
  movel([0.423322, -1.407302, -2.551374, -0.753713, 1.570796, 1.994118],accel_mss,speed_ms,0,blend_radius_m)
  movel([0.424496, -1.407939, -2.550899, -0.753551, 1.570796, 1.995293],accel_mss,speed_ms,0,blend_radius_m)
  movel([0.425844, -1.408177, -2.550722, -0.753490, 1.570796, 1.996641],accel_mss,speed_ms,0,blend_radius_m)
  movel([0.427662, -1.407960, -2.550884, -0.753545, 1.570796, 1.998458],accel_mss,speed_ms,0,blend_radius_m)
  movel([0.428488, -1.407649, -2.551116, -0.753624, 1.570796, 1.999285],accel_mss,speed_ms,0,blend_radius_m)
  movel([0.429264, -1.407205, -2.551446, -0.753737, 1.570796, 2.000060],accel_mss,speed_ms,0,blend_radius_m)
  movel([0.430547, -1.406086, -2.552279, -0.754024, 1.570796, 2.001343],accel_mss,speed_ms,0,blend_radius_m)
  movel([0.431417, -1.404767, -2.553258, -0.754364, 1.570796, 2.002214],accel_mss,speed_ms,0,blend_radius_m)
  movel([0.431738, -1.403866, -2.553925, -0.754598, 1.570796, 2.002535],accel_mss,speed_ms,0,blend_radius_m)
  movel([0.431756, -1.403191, -2.554424, -0.754773, 1.570796, 2.002553],accel_mss,speed_ms,0,blend_radius_m)
  movel([0.431510, -1.402769, -2.554736, -0.754884, 1.570796, 2.002306],accel_mss,speed_ms,0,blend_radius_m)
  movel([0.431043, -1.402615, -2.554850, -0.754924, 1.570796, 2.001840],accel_mss,speed_ms,0,blend_radius_m)
  movel([0.430110, -1.402919, -2.554626, -0.754845, 1.570796, 2.000906],accel_mss,speed_ms,0,blend_radius_m)
  movel([0.429188, -1.403285, -2.554355, -0.754749, 1.570796, 1.999985],accel_mss,speed_ms,0,blend_radius_m)
  movel([0.428133, -1.403402, -2.554269, -0.754719, 1.570796, 1.998930],accel_mss,speed_ms,0,blend_radius_m)
  movel([0.427069, -1.403144, -2.554459, -0.754786, 1.570796, 1.997865],accel_mss,speed_ms,0,blend_radius_m)
  movel([0.426515, -1.402437, -2.554981, -0.754971, 1.570796, 1.997312],accel_mss,speed_ms,0,blend_radius_m)
  movel([0.426435, -1.401422, -2.555729, -0.755238, 1.570796, 1.997232],accel_mss,speed_ms,0,blend_radius_m)
  movel([0.426796, -1.400238, -2.556600, -0.755551, 1.570796, 1.997592],accel_mss,speed_ms,0,blend_radius_m)
  movel([0.427523, -1.399062, -2.557463, -0.755864, 1.570796, 1.998320],accel_mss,speed_ms,0,blend_radius_m)
  movel([0.428532, -1.398067, -2.558191, -0.756131, 1.570796, 1.999328],accel_mss,speed_ms,0,blend_radius_m)
  movel([0.429727, -1.397396, -2.558682, -0.756311, 1.570796, 2.000524],accel_mss,speed_ms,0,blend_radius_m)
  movel([0.431011, -1.397195, -2.558829, -0.756365, 1.570796, 2.001808],accel_mss,speed_ms,0,blend_radius_m)
  movel([0.431985, -1.397355, -2.558712, -0.756322, 1.570796, 2.002781],accel_mss,speed_ms,0,blend_radius_m)
  movel([0.432705, -1.397780, -2.558401, -0.756208, 1.570796, 2.003502],accel_mss,speed_ms,0,blend_radius_m)
  movel([0.433176, -1.398467, -2.557899, -0.756023, 1.570796, 2.003973],accel_mss,speed_ms,0,blend_radius_m)
  movel([0.433392, -1.399418, -2.557202, -0.755769, 1.570796, 2.004188],accel_mss,speed_ms,0,blend_radius_m)
  movel([0.433378, -1.400563, -2.556361, -0.755465, 1.570796, 2.004174],accel_mss,speed_ms,0,blend_radius_m)
  movel([0.433152, -1.401841, -2.555420, -0.755127, 1.570796, 2.003949],accel_mss,speed_ms,0,blend_radius_m)
  movel([0.432073, -1.404786, -2.553244, -0.754359, 1.570796, 2.002870],accel_mss,speed_ms,0,blend_radius_m)
  movel([0.431091, -1.406675, -2.551841, -0.753873, 1.570796, 2.001887],accel_mss,speed_ms,0,blend_radius_m)
  movel([0.429960, -1.408447, -2.550520, -0.753422, 1.570796, 2.000756],accel_mss,speed_ms,0,blend_radius_m)
  movel([0.428685, -1.410108, -2.549278, -0.753003, 1.570796, 1.999481],accel_mss,speed_ms,0,blend_radius_m)
  movel([0.427260, -1.411655, -2.548118, -0.752617, 1.570796, 1.998056],accel_mss,speed_ms,0,blend_radius_m)
  movel([0.425714, -1.412954, -2.547140, -0.752295, 1.570796, 1.996510],accel_mss,speed_ms,0,blend_radius_m)
  movel([0.424071, -1.413866, -2.546453, -0.752071, 1.570796, 1.994867],accel_mss,speed_ms,0,blend_radius_m)
  movel([0.422329, -1.414394, -2.546054, -0.751941, 1.570796, 1.993125],accel_mss,speed_ms,0,blend_radius_m)
  movel([0.420484, -1.414542, -2.545942, -0.751905, 1.570796, 1.991281],accel_mss,speed_ms,0,blend_radius_m)
  movel([0.418943, -1.414337, -2.546097, -0.751955, 1.570796, 1.989740],accel_mss,speed_ms,0,blend_radius_m)
  movel([0.417669, -1.413798, -2.546504, -0.752087, 1.570796, 1.988465],accel_mss,speed_ms,0,blend_radius_m)
  movel([0.416628, -1.413010, -2.547098, -0.752281, 1.570796, 1.987424],accel_mss,speed_ms,0,blend_radius_m)
  movel([0.415791, -1.412067, -2.547808, -0.752514, 1.570796, 1.986587],accel_mss,speed_ms,0,blend_radius_m)
  movel([0.414190, -1.409372, -2.549829, -0.753188, 1.570796, 1.984986],accel_mss,speed_ms,0,blend_radius_m)
  movel([0.412653, -1.406837, -2.551721, -0.753832, 1.570796, 1.983449],accel_mss,speed_ms,0,blend_radius_m)
  movel([0.411886, -1.405968, -2.552367, -0.754054, 1.570796, 1.982682],accel_mss,speed_ms,0,blend_radius_m)
  movel([0.410949, -1.405252, -2.552898, -0.754238, 1.570796, 1.981745],accel_mss,speed_ms,0,blend_radius_m)
  movel([0.409814, -1.404771, -2.553255, -0.754363, 1.570796, 1.980610],accel_mss,speed_ms,0,blend_radius_m)
  movel([0.408469, -1.404603, -2.553380, -0.754406, 1.570796, 1.979265],accel_mss,speed_ms,0,blend_radius_m)
  movel([0.408146, -1.405334, -2.552838, -0.754218, 1.570796, 1.978942],accel_mss,speed_ms,0,blend_radius_m)
  movel([0.407355, -1.407354, -2.551336, -0.753700, 1.570796, 1.978152],accel_mss,speed_ms,0,blend_radius_m)
  movel([0.406880, -1.409123, -2.550015, -0.753251, 1.570796, 1.977676],accel_mss,speed_ms,0,blend_radius_m)
  movel([0.406719, -1.410644, -2.548876, -0.752869, 1.570796, 1.977515],accel_mss,speed_ms,0,blend_radius_m)
  movel([0.406870, -1.411917, -2.547920, -0.752551, 1.570796, 1.977667],accel_mss,speed_ms,0,blend_radius_m)
  movel([0.407293, -1.412956, -2.547139, -0.752294, 1.570796, 1.978089],accel_mss,speed_ms,0,blend_radius_m)
  movel([0.407940, -1.413775, -2.546521, -0.752093, 1.570796, 1.978736],accel_mss,speed_ms,0,blend_radius_m)
  movel([0.408816, -1.414378, -2.546066, -0.751945, 1.570796, 1.979612],accel_mss,speed_ms,0,blend_radius_m)
  movel([0.409919, -1.414761, -2.545776, -0.751852, 1.570796, 1.980715],accel_mss,speed_ms,0,blend_radius_m)
  movel([0.403355, -1.414702, -2.545821, -0.751866, 1.570796, 1.974151],accel_mss,speed_ms,0,blend_radius_m)
  movel([0.411975, -1.395197, -2.560284, -0.756907, 1.570796, 1.982772],accel_mss,speed_ms,0,blend_radius_m)
  movel([0.412645, -1.395201, -2.560281, -0.756906, 1.570796, 1.983441],accel_mss,speed_ms,0,blend_radius_m)
  speed_ms = 0.003
  movel([0.412645, -1.388740, -2.557323, -0.766326, 1.570796, 1.983441],accel_mss,speed_ms,0,blend_radius_m)
  speed_ms = 0.03
  movel([0.412645, -1.363842, -2.545198, -0.803350, 1.570796, 1.983441],accel_mss,speed_ms,0,blend_radius_m)
  #M_RunCode9
  movel([0.406400, -1.386317, -2.529254, -0.796817, 1.570796, 1.977196],accel_mss,speed_ms,0,blend_radius_m)
  #M_RunCode3
  movel([0.406400, -1.410785, -2.541097, -0.760508, 1.570796, 1.977196],accel_mss,speed_ms,0,blend_radius_m)
  speed_ms = 0.003
  movel([0.406400, -1.417125, -2.543985, -0.751279, 1.570796, 1.977196],accel_mss,speed_ms,0,blend_radius_m)
  speed_ms = 0.007
  movel([0.407465, -1.417363, -2.543804, -0.751222, 1.570796, 1.978262],accel_mss,speed_ms,0,blend_radius_m)
  movel([0.408048, -1.418042, -2.543288, -0.751059, 1.570796, 1.978844],accel_mss,speed_ms,0,blend_radius_m)
  movel([0.408163, -1.419027, -2.542537, -0.750824, 1.570796, 1.978960],accel_mss,speed_ms,0,blend_radius_m)
  movel([0.407837, -1.420174, -2.541662, -0.750553, 1.570796, 1.978633],accel_mss,speed_ms,0,blend_radius_m)
  movel([0.407147, -1.421313, -2.540791, -0.750285, 1.570796, 1.977944],accel_mss,speed_ms,0,blend_radius_m)
  movel([0.406168, -1.422279, -2.540051, -0.750060, 1.570796, 1.976964],accel_mss,speed_ms,0,blend_radius_m)
  movel([0.404997, -1.422935, -2.539547, -0.749907, 1.570796, 1.975794],accel_mss,speed_ms,0,blend_radius_m)
  movel([0.403741, -1.423144, -2.539386, -0.749859, 1.570796, 1.974538],accel_mss,speed_ms,0,blend_radius_m)
  movel([0.402826, -1.422997, -2.539499, -0.749893, 1.570796, 1.973622],accel_mss,speed_ms,0,blend_radius_m)
  movel([0.402259, -1.422617, -2.539791, -0.749981, 1.570796, 1.973055],accel_mss,speed_ms,0,blend_radius_m)
  movel([0.401621, -1.422296, -2.540038, -0.750056, 1.570796, 1.972418],accel_mss,speed_ms,0,blend_radius_m)
  movel([0.401037, -1.422430, -2.539934, -0.750024, 1.570796, 1.971834],accel_mss,speed_ms,0,blend_radius_m)
  movel([0.400423, -1.422843, -2.539618, -0.749929, 1.570796, 1.971219],accel_mss,speed_ms,0,blend_radius_m)
  movel([0.399871, -1.423441, -2.539158, -0.749790, 1.570796, 1.970667],accel_mss,speed_ms,0,blend_radius_m)
  movel([0.399469, -1.424139, -2.538621, -0.749629, 1.570796, 1.970265],accel_mss,speed_ms,0,blend_radius_m)
  movel([0.399162, -1.425063, -2.537909, -0.749418, 1.570796, 1.969959],accel_mss,speed_ms,0,blend_radius_m)
  movel([0.399089, -1.425906, -2.537258, -0.749225, 1.570796, 1.969885],accel_mss,speed_ms,0,blend_radius_m)
  movel([0.399247, -1.426667, -2.536670, -0.749053, 1.570796, 1.970043],accel_mss,speed_ms,0,blend_radius_m)
  movel([0.399633, -1.427350, -2.536140, -0.748899, 1.570796, 1.970429],accel_mss,speed_ms,0,blend_radius_m)
  movel([0.400227, -1.427912, -2.535705, -0.748772, 1.570796, 1.971023],accel_mss,speed_ms,0,blend_radius_m)
  movel([0.401003, -1.428317, -2.535390, -0.748682, 1.570796, 1.971800],accel_mss,speed_ms,0,blend_radius_m)
  movel([0.401961, -1.428566, -2.535197, -0.748626, 1.570796, 1.972758],accel_mss,speed_ms,0,blend_radius_m)
  movel([0.403101, -1.428658, -2.535125, -0.748605, 1.570796, 1.973898],accel_mss,speed_ms,0,blend_radius_m)
  movel([0.405186, -1.428400, -2.535326, -0.748663, 1.570796, 1.975982],accel_mss,speed_ms,0,blend_radius_m)
  movel([0.407320, -1.427574, -2.535967, -0.748848, 1.570796, 1.978116],accel_mss,speed_ms,0,blend_radius_m)
  movel([0.408394, -1.426941, -2.536457, -0.748991, 1.570796, 1.979190],accel_mss,speed_ms,0,blend_radius_m)
  movel([0.409447, -1.426161, -2.537060, -0.749167, 1.570796, 1.980243],accel_mss,speed_ms,0,blend_radius_m)
  movel([0.411502, -1.424141, -2.538619, -0.749629, 1.570796, 1.982298],accel_mss,speed_ms,0,blend_radius_m)
  movel([0.413409, -1.421538, -2.540619, -0.750233, 1.570796, 1.984205],accel_mss,speed_ms,0,blend_radius_m)
  movel([0.415084, -1.418369, -2.543039, -0.750981, 1.570796, 1.985881],accel_mss,speed_ms,0,blend_radius_m)
  movel([0.425033, -1.418605, -2.542859, -0.750925, 1.570796, 1.995830],accel_mss,speed_ms,0,blend_radius_m)
  movel([0.418518, -1.432773, -2.531916, -0.747700, 1.570796, 1.989314],accel_mss,speed_ms,0,blend_radius_m)
  movel([0.412120, -1.432614, -2.532040, -0.747734, 1.570796, 1.982916],accel_mss,speed_ms,0,blend_radius_m)
  movel([0.413891, -1.432114, -2.532432, -0.747843, 1.570796, 1.984687],accel_mss,speed_ms,0,blend_radius_m)
  movel([0.415728, -1.431165, -2.533173, -0.748051, 1.570796, 1.986525],accel_mss,speed_ms,0,blend_radius_m)
  movel([0.417541, -1.429812, -2.534228, -0.748349, 1.570796, 1.988337],accel_mss,speed_ms,0,blend_radius_m)
  movel([0.419237, -1.428099, -2.535559, -0.748730, 1.570796, 1.990033],accel_mss,speed_ms,0,blend_radius_m)
  movel([0.420743, -1.426078, -2.537125, -0.749186, 1.570796, 1.991539],accel_mss,speed_ms,0,blend_radius_m)
  movel([0.421981, -1.423804, -2.538878, -0.749706, 1.570796, 1.992777],accel_mss,speed_ms,0,blend_radius_m)
  movel([0.414673, -1.423628, -2.539014, -0.749747, 1.570796, 1.985469],accel_mss,speed_ms,0,blend_radius_m)
  movel([0.413202, -1.426433, -2.536850, -0.749106, 1.570796, 1.983998],accel_mss,speed_ms,0,blend_radius_m)
  movel([0.411390, -1.429102, -2.534780, -0.748507, 1.570796, 1.982186],accel_mss,speed_ms,0,blend_radius_m)
  movel([0.409295, -1.431455, -2.532947, -0.747987, 1.570796, 1.980092],accel_mss,speed_ms,0,blend_radius_m)
  movel([0.408161, -1.432447, -2.532171, -0.747771, 1.570796, 1.978958],accel_mss,speed_ms,0,blend_radius_m)
  movel([0.406973, -1.433318, -2.531489, -0.747582, 1.570796, 1.977769],accel_mss,speed_ms,0,blend_radius_m)
  movel([0.405742, -1.434024, -2.530935, -0.747430, 1.570796, 1.976539],accel_mss,speed_ms,0,blend_radius_m)
  movel([0.404493, -1.434523, -2.530544, -0.747323, 1.570796, 1.975289],accel_mss,speed_ms,0,blend_radius_m)
  movel([0.403220, -1.434816, -2.530313, -0.747260, 1.570796, 1.974017],accel_mss,speed_ms,0,blend_radius_m)
  movel([0.401929, -1.434901, -2.530246, -0.747242, 1.570796, 1.972725],accel_mss,speed_ms,0,blend_radius_m)
  movel([0.400722, -1.434790, -2.530333, -0.747265, 1.570796, 1.971518],accel_mss,speed_ms,0,blend_radius_m)
  movel([0.399703, -1.434491, -2.530568, -0.747329, 1.570796, 1.970499],accel_mss,speed_ms,0,blend_radius_m)
  movel([0.398876, -1.434002, -2.530952, -0.747434, 1.570796, 1.969672],accel_mss,speed_ms,0,blend_radius_m)
  movel([0.398239, -1.433325, -2.531484, -0.747580, 1.570796, 1.969036],accel_mss,speed_ms,0,blend_radius_m)
  movel([0.397478, -1.431573, -2.532855, -0.747961, 1.570796, 1.968274],accel_mss,speed_ms,0,blend_radius_m)
  movel([0.397353, -1.429412, -2.534539, -0.748438, 1.570796, 1.968149],accel_mss,speed_ms,0,blend_radius_m)
  movel([0.397775, -1.427007, -2.536406, -0.748976, 1.570796, 1.968571],accel_mss,speed_ms,0,blend_radius_m)
  movel([0.398644, -1.424530, -2.538319, -0.749539, 1.570796, 1.969441],accel_mss,speed_ms,0,blend_radius_m)
  movel([0.399519, -1.422827, -2.539630, -0.749932, 1.570796, 1.970316],accel_mss,speed_ms,0,blend_radius_m)
  movel([0.400673, -1.421101, -2.540953, -0.750335, 1.570796, 1.971469],accel_mss,speed_ms,0,blend_radius_m)
  movel([0.402021, -1.419516, -2.542165, -0.750709, 1.570796, 1.972817],accel_mss,speed_ms,0,blend_radius_m)
  movel([0.403484, -1.418239, -2.543137, -0.751012, 1.570796, 1.974280],accel_mss,speed_ms,0,blend_radius_m)
  movel([0.404974, -1.417397, -2.543778, -0.751214, 1.570796, 1.975770],accel_mss,speed_ms,0,blend_radius_m)
  movel([0.406400, -1.417125, -2.543985, -0.751279, 1.570796, 1.977196],accel_mss,speed_ms,0,blend_radius_m)
  speed_ms = 0.003
  movel([0.406400, -1.410785, -2.541097, -0.760508, 1.570796, 1.977196],accel_mss,speed_ms,0,blend_radius_m)
  speed_ms = 0.03
  movel([0.406400, -1.386317, -2.529254, -0.796817, 1.570796, 1.977196],accel_mss,speed_ms,0,blend_radius_m)
  #M_RunCode9
  movel([0.492309, -1.304268, -2.584161, -0.823959, 1.570796, 2.063105],accel_mss,speed_ms,0,blend_radius_m)
  #M_RunCode3
  movel([0.492309, -1.330216, -2.597053, -0.785121, 1.570796, 2.063105],accel_mss,speed_ms,0,blend_radius_m)
  speed_ms = 0.003
  movel([0.492309, -1.336975, -2.600204, -0.775209, 1.570796, 2.063105],accel_mss,speed_ms,0,blend_radius_m)
  speed_ms = 0.007
  movel([0.492396, -1.336918, -2.600241, -0.775230, 1.570796, 2.063192],accel_mss,speed_ms,0,blend_radius_m)
  movel([0.492309, -1.336975, -2.600204, -0.775209, 1.570796, 2.063105],accel_mss,speed_ms,0,blend_radius_m)
  speed_ms = 0.003
  movel([0.492309, -1.330216, -2.597053, -0.785121, 1.570796, 2.063105],accel_mss,speed_ms,0,blend_radius_m)
  speed_ms = 0.03
  movel([0.492309, -1.304268, -2.584161, -0.823959, 1.570796, 2.063105],accel_mss,speed_ms,0,blend_radius_m)
  #M_RunCode9
  movel([0.469500, -1.315047, -2.577456, -0.819886, 1.570796, 2.040297],accel_mss,speed_ms,0,blend_radius_m)
  #M_RunCode3
  movel([0.469500, -1.340816, -2.590208, -0.781365, 1.570796, 2.040297],accel_mss,speed_ms,0,blend_radius_m)
  speed_ms = 0.003
  movel([0.469500, -1.347524, -2.593324, -0.771541, 1.570796, 2.040297],accel_mss,speed_ms,0,blend_radius_m)
  speed_ms = 0.007
  movel([0.469474, -1.348724, -2.592531, -0.771133, 1.570796, 2.040271],accel_mss,speed_ms,0,blend_radius_m)
  movel([0.469105, -1.350166, -2.591577, -0.770646, 1.570796, 2.039902],accel_mss,speed_ms,0,blend_radius_m)
  movel([0.468017, -1.352314, -2.590149, -0.769926, 1.570796, 2.038814],accel_mss,speed_ms,0,blend_radius_m)
  movel([0.466438, -1.354171, -2.588910, -0.769308, 1.570796, 2.037234],accel_mss,speed_ms,0,blend_radius_m)
  movel([0.464459, -1.355721, -2.587872, -0.768796, 1.570796, 2.035256],accel_mss,speed_ms,0,blend_radius_m)
  movel([0.462181, -1.356944, -2.587050, -0.768395, 1.570796, 2.032977],accel_mss,speed_ms,0,blend_radius_m)
  movel([0.459591, -1.357798, -2.586475, -0.768116, 1.570796, 2.030388],accel_mss,speed_ms,0,blend_radius_m)
  movel([0.457486, -1.357931, -2.586385, -0.768072, 1.570796, 2.028282],accel_mss,speed_ms,0,blend_radius_m)
  movel([0.455825, -1.357452, -2.586708, -0.768229, 1.570796, 2.026621],accel_mss,speed_ms,0,blend_radius_m)
  movel([0.454572, -1.356458, -2.587376, -0.768554, 1.570796, 2.025369],accel_mss,speed_ms,0,blend_radius_m)
  movel([0.453687, -1.355057, -2.588317, -0.769015, 1.570796, 2.024483],accel_mss,speed_ms,0,blend_radius_m)
  movel([0.453136, -1.353349, -2.589459, -0.769581, 1.570796, 2.023932],accel_mss,speed_ms,0,blend_radius_m)
  movel([0.452883, -1.351439, -2.590731, -0.770219, 1.570796, 2.023680],accel_mss,speed_ms,0,blend_radius_m)
  movel([0.452896, -1.349430, -2.592065, -0.770895, 1.570796, 2.023692],accel_mss,speed_ms,0,blend_radius_m)
  movel([0.455382, -1.347696, -2.593210, -0.771482, 1.570796, 2.026178],accel_mss,speed_ms,0,blend_radius_m)
  movel([0.458299, -1.346270, -2.594150, -0.771969, 1.570796, 2.029096],accel_mss,speed_ms,0,blend_radius_m)
  movel([0.461367, -1.345261, -2.594813, -0.772315, 1.570796, 2.032163],accel_mss,speed_ms,0,blend_radius_m)
  movel([0.464301, -1.344777, -2.595131, -0.772482, 1.570796, 2.035097],accel_mss,speed_ms,0,blend_radius_m)
  movel([0.466823, -1.344925, -2.595034, -0.772431, 1.570796, 2.037620],accel_mss,speed_ms,0,blend_radius_m)
  movel([0.467840, -1.345270, -2.594807, -0.772312, 1.570796, 2.038636],accel_mss,speed_ms,0,blend_radius_m)
  movel([0.468649, -1.345809, -2.594453, -0.772127, 1.570796, 2.039445],accel_mss,speed_ms,0,blend_radius_m)
  movel([0.469213, -1.346556, -2.593962, -0.771871, 1.570796, 2.040009],accel_mss,speed_ms,0,blend_radius_m)
  movel([0.469500, -1.347524, -2.593324, -0.771541, 1.570796, 2.040297],accel_mss,speed_ms,0,blend_radius_m)
  speed_ms = 0.003
  movel([0.469500, -1.340816, -2.590208, -0.781365, 1.570796, 2.040297],accel_mss,speed_ms,0,blend_radius_m)
  speed_ms = 0.03
  movel([0.469500, -1.315047, -2.577456, -0.819886, 1.570796, 2.040297],accel_mss,speed_ms,0,blend_radius_m)
  #M_RunCode9
  movel([0.530434, -1.300426, -2.586516, -0.825448, 1.570796, 2.101230],accel_mss,speed_ms,0,blend_radius_m)
  #M_RunCode3
  movel([0.530434, -1.326435, -2.599457, -0.786496, 1.570796, 2.101230],accel_mss,speed_ms,0,blend_radius_m)
  speed_ms = 0.003
  movel([0.530434, -1.333213, -2.602622, -0.776555, 1.570796, 2.101230],accel_mss,speed_ms,0,blend_radius_m)
  speed_ms = 0.007
  movel([0.531089, -1.331788, -2.603532, -0.777069, 1.570796, 2.101886],accel_mss,speed_ms,0,blend_radius_m)
  movel([0.531935, -1.330340, -2.604454, -0.777595, 1.570796, 2.102732],accel_mss,speed_ms,0,blend_radius_m)
  movel([0.532293, -1.330582, -2.604300, -0.777506, 1.570796, 2.103089],accel_mss,speed_ms,0,blend_radius_m)
  movel([0.532242, -1.331062, -2.603995, -0.777332, 1.570796, 2.103038],accel_mss,speed_ms,0,blend_radius_m)
  movel([0.532223, -1.331603, -2.603650, -0.777136, 1.570796, 2.103020],accel_mss,speed_ms,0,blend_radius_m)
  movel([0.532677, -1.332026, -2.603380, -0.776983, 1.570796, 2.103473],accel_mss,speed_ms,0,blend_radius_m)
  movel([0.533455, -1.332142, -2.603306, -0.776941, 1.570796, 2.104251],accel_mss,speed_ms,0,blend_radius_m)
  movel([0.534342, -1.332066, -2.603355, -0.776968, 1.570796, 2.105138],accel_mss,speed_ms,0,blend_radius_m)
  movel([0.535593, -1.331910, -2.603454, -0.777025, 1.570796, 2.106390],accel_mss,speed_ms,0,blend_radius_m)
  movel([0.536736, -1.330110, -2.604600, -0.777678, 1.570796, 2.107533],accel_mss,speed_ms,0,blend_radius_m)
  movel([0.537276, -1.328570, -2.605578, -0.778241, 1.570796, 2.108072],accel_mss,speed_ms,0,blend_radius_m)
  movel([0.537238, -1.327949, -2.605971, -0.778469, 1.570796, 2.108034],accel_mss,speed_ms,0,blend_radius_m)
  movel([0.536958, -1.327456, -2.606283, -0.778650, 1.570796, 2.107755],accel_mss,speed_ms,0,blend_radius_m)
  movel([0.536401, -1.327111, -2.606501, -0.778777, 1.570796, 2.107197],accel_mss,speed_ms,0,blend_radius_m)
  movel([0.535536, -1.326937, -2.606611, -0.778841, 1.570796, 2.106332],accel_mss,speed_ms,0,blend_radius_m)
  movel([0.536562, -1.326099, -2.607140, -0.779150, 1.570796, 2.107358],accel_mss,speed_ms,0,blend_radius_m)
  movel([0.537493, -1.325468, -2.607537, -0.779384, 1.570796, 2.108290],accel_mss,speed_ms,0,blend_radius_m)
  movel([0.537872, -1.325336, -2.607620, -0.779433, 1.570796, 2.108668],accel_mss,speed_ms,0,blend_radius_m)
  movel([0.538164, -1.325378, -2.607594, -0.779417, 1.570796, 2.108960],accel_mss,speed_ms,0,blend_radius_m)
  movel([0.538409, -1.326155, -2.607104, -0.779130, 1.570796, 2.109205],accel_mss,speed_ms,0,blend_radius_m)
  movel([0.538144, -1.328153, -2.605842, -0.778394, 1.570796, 2.108940],accel_mss,speed_ms,0,blend_radius_m)
  movel([0.537378, -1.330295, -2.604483, -0.777611, 1.570796, 2.108174],accel_mss,speed_ms,0,blend_radius_m)
  movel([0.536791, -1.331316, -2.603833, -0.777240, 1.570796, 2.107587],accel_mss,speed_ms,0,blend_radius_m)
  movel([0.536052, -1.332251, -2.603236, -0.776901, 1.570796, 2.106849],accel_mss,speed_ms,0,blend_radius_m)
  movel([0.535159, -1.333057, -2.602722, -0.776611, 1.570796, 2.105955],accel_mss,speed_ms,0,blend_radius_m)
  movel([0.534100, -1.333693, -2.602314, -0.776382, 1.570796, 2.104897],accel_mss,speed_ms,0,blend_radius_m)
  movel([0.534211, -1.332459, -2.603104, -0.776826, 1.570796, 2.105008],accel_mss,speed_ms,0,blend_radius_m)
  movel([0.530368, -1.335772, -2.600979, -0.775637, 1.570796, 2.101165],accel_mss,speed_ms,0,blend_radius_m)
  movel([0.530138, -1.334560, -2.601758, -0.776071, 1.570796, 2.100934],accel_mss,speed_ms,0,blend_radius_m)
  movel([0.530434, -1.333213, -2.602622, -0.776555, 1.570796, 2.101230],accel_mss,speed_ms,0,blend_radius_m)
  speed_ms = 0.003
  movel([0.530434, -1.326435, -2.599457, -0.786496, 1.570796, 2.101230],accel_mss,speed_ms,0,blend_radius_m)
  speed_ms = 0.03
  movel([0.530434, -1.300426, -2.586516, -0.825448, 1.570796, 2.101230],accel_mss,speed_ms,0,blend_radius_m)
  #M_RunCode9
  movel([0.547267, -1.261948, -2.609078, -0.841364, 1.570796, 2.118063],accel_mss,speed_ms,0,blend_radius_m)
  #M_RunCode3
  movel([0.547267, -1.288536, -2.622525, -0.801328, 1.570796, 2.118063],accel_mss,speed_ms,0,blend_radius_m)
  speed_ms = 0.003
  movel([0.547267, -1.295484, -2.625817, -0.791088, 1.570796, 2.118063],accel_mss,speed_ms,0,blend_radius_m)
  speed_ms = 0.007
  movel([0.545499, -1.295503, -2.625806, -0.791080, 1.570796, 2.116295],accel_mss,speed_ms,0,blend_radius_m)
  movel([0.543826, -1.295292, -2.625930, -0.791167, 1.570796, 2.114622],accel_mss,speed_ms,0,blend_radius_m)
  movel([0.542273, -1.294844, -2.626194, -0.791350, 1.570796, 2.113069],accel_mss,speed_ms,0,blend_radius_m)
  movel([0.540868, -1.294147, -2.626605, -0.791637, 1.570796, 2.111664],accel_mss,speed_ms,0,blend_radius_m)
  movel([0.539637, -1.293197, -2.627164, -0.792029, 1.570796, 2.110433],accel_mss,speed_ms,0,blend_radius_m)
  movel([0.539192, -1.292496, -2.627575, -0.792318, 1.570796, 2.109988],accel_mss,speed_ms,0,blend_radius_m)
  movel([0.538882, -1.291626, -2.628084, -0.792679, 1.570796, 2.109678],accel_mss,speed_ms,0,blend_radius_m)
  movel([0.538600, -1.290849, -2.628538, -0.793002, 1.570796, 2.109396],accel_mss,speed_ms,0,blend_radius_m)
  movel([0.538231, -1.290425, -2.628786, -0.793178, 1.570796, 2.109027],accel_mss,speed_ms,0,blend_radius_m)
  movel([0.537072, -1.290379, -2.628813, -0.793197, 1.570796, 2.107869],accel_mss,speed_ms,0,blend_radius_m)
  movel([0.535335, -1.290591, -2.628689, -0.793109, 1.570796, 2.106131],accel_mss,speed_ms,0,blend_radius_m)
  movel([0.533504, -1.290841, -2.628543, -0.793005, 1.570796, 2.104300],accel_mss,speed_ms,0,blend_radius_m)
  movel([0.532068, -1.290903, -2.628507, -0.792979, 1.570796, 2.102864],accel_mss,speed_ms,0,blend_radius_m)
  movel([0.529688, -1.290429, -2.628784, -0.793176, 1.570796, 2.100484],accel_mss,speed_ms,0,blend_radius_m)
  movel([0.527892, -1.289567, -2.629286, -0.793535, 1.570796, 2.098688],accel_mss,speed_ms,0,blend_radius_m)
  movel([0.526627, -1.288358, -2.629989, -0.794041, 1.570796, 2.097423],accel_mss,speed_ms,0,blend_radius_m)
  movel([0.525845, -1.286838, -2.630871, -0.794680, 1.570796, 2.096641],accel_mss,speed_ms,0,blend_radius_m)
  movel([0.525498, -1.285041, -2.631910, -0.795438, 1.570796, 2.096295],accel_mss,speed_ms,0,blend_radius_m)
  movel([0.525534, -1.283007, -2.633080, -0.796301, 1.570796, 2.096331],accel_mss,speed_ms,0,blend_radius_m)
  movel([0.525907, -1.280776, -2.634358, -0.797254, 1.570796, 2.096703],accel_mss,speed_ms,0,blend_radius_m)
  movel([0.526562, -1.278382, -2.635723, -0.798284, 1.570796, 2.097358],accel_mss,speed_ms,0,blend_radius_m)
  movel([0.528525, -1.273279, -2.638607, -0.800503, 1.570796, 2.099321],accel_mss,speed_ms,0,blend_radius_m)
  movel([0.531020, -1.268018, -2.641547, -0.802824, 1.570796, 2.101816],accel_mss,speed_ms,0,blend_radius_m)
  movel([0.535903, -1.258402, -2.646832, -0.807155, 1.570796, 2.106699],accel_mss,speed_ms,0,blend_radius_m)
  movel([0.537738, -1.254140, -2.649139, -0.809110, 1.570796, 2.108534],accel_mss,speed_ms,0,blend_radius_m)
  movel([0.539517, -1.249200, -2.651785, -0.811404, 1.570796, 2.110313],accel_mss,speed_ms,0,blend_radius_m)
  movel([0.541129, -1.243838, -2.654624, -0.813927, 1.570796, 2.111926],accel_mss,speed_ms,0,blend_radius_m)
  movel([0.542464, -1.238310, -2.657516, -0.816563, 1.570796, 2.113260],accel_mss,speed_ms,0,blend_radius_m)
  movel([0.543395, -1.232890, -2.660316, -0.819183, 1.570796, 2.114192],accel_mss,speed_ms,0,blend_radius_m)
  movel([0.543802, -1.227852, -2.662888, -0.821649, 1.570796, 2.114599],accel_mss,speed_ms,0,blend_radius_m)
  movel([0.543559, -1.223489, -2.665092, -0.823808, 1.570796, 2.114355],accel_mss,speed_ms,0,blend_radius_m)
  movel([0.543154, -1.221653, -2.666013, -0.824723, 1.570796, 2.113950],accel_mss,speed_ms,0,blend_radius_m)
  movel([0.542538, -1.220095, -2.666791, -0.825503, 1.570796, 2.113335],accel_mss,speed_ms,0,blend_radius_m)
  movel([0.541649, -1.218693, -2.667489, -0.826207, 1.570796, 2.112445],accel_mss,speed_ms,0,blend_radius_m)
  movel([0.540377, -1.217258, -2.668201, -0.826929, 1.570796, 2.111173],accel_mss,speed_ms,0,blend_radius_m)
  movel([0.538740, -1.215933, -2.668857, -0.827599, 1.570796, 2.109537],accel_mss,speed_ms,0,blend_radius_m)
  movel([0.536764, -1.214856, -2.669388, -0.828144, 1.570796, 2.107560],accel_mss,speed_ms,0,blend_radius_m)
  movel([0.534467, -1.214178, -2.669722, -0.828489, 1.570796, 2.105263],accel_mss,speed_ms,0,blend_radius_m)
  movel([0.531876, -1.214037, -2.669792, -0.828560, 1.570796, 2.102673],accel_mss,speed_ms,0,blend_radius_m)
  movel([0.529019, -1.214575, -2.669527, -0.828287, 1.570796, 2.099815],accel_mss,speed_ms,0,blend_radius_m)
  movel([0.527498, -1.215144, -2.669246, -0.827999, 1.570796, 2.098294],accel_mss,speed_ms,0,blend_radius_m)
  movel([0.525923, -1.215932, -2.668858, -0.827600, 1.570796, 2.096719],accel_mss,speed_ms,0,blend_radius_m)
  movel([0.523569, -1.217549, -2.668057, -0.826783, 1.570796, 2.094365],accel_mss,speed_ms,0,blend_radius_m)
  movel([0.521715, -1.219421, -2.667127, -0.825841, 1.570796, 2.092511],accel_mss,speed_ms,0,blend_radius_m)
  movel([0.520317, -1.221504, -2.666087, -0.824798, 1.570796, 2.091114],accel_mss,speed_ms,0,blend_radius_m)
  movel([0.519329, -1.223761, -2.664955, -0.823673, 1.570796, 2.090125],accel_mss,speed_ms,0,blend_radius_m)
  movel([0.518708, -1.226153, -2.663749, -0.822487, 1.570796, 2.089504],accel_mss,speed_ms,0,blend_radius_m)
  movel([0.518400, -1.228649, -2.662483, -0.821257, 1.570796, 2.089196],accel_mss,speed_ms,0,blend_radius_m)
  movel([0.518359, -1.231209, -2.661177, -0.820003, 1.570796, 2.089155],accel_mss,speed_ms,0,blend_radius_m)
  movel([0.518541, -1.233802, -2.659847, -0.818740, 1.570796, 2.089338],accel_mss,speed_ms,0,blend_radius_m)
  movel([0.519379, -1.238946, -2.657185, -0.816258, 1.570796, 2.090176],accel_mss,speed_ms,0,blend_radius_m)
  movel([0.520552, -1.243813, -2.654638, -0.813939, 1.570796, 2.091349],accel_mss,speed_ms,0,blend_radius_m)
  movel([0.521703, -1.248132, -2.652353, -0.811904, 1.570796, 2.092500],accel_mss,speed_ms,0,blend_radius_m)
  movel([0.522479, -1.251644, -2.650480, -0.810266, 1.570796, 2.093275],accel_mss,speed_ms,0,blend_radius_m)
  movel([0.523939, -1.260309, -2.645793, -0.806287, 1.570796, 2.094736],accel_mss,speed_ms,0,blend_radius_m)
  movel([0.524584, -1.264978, -2.643230, -0.804181, 1.570796, 2.095380],accel_mss,speed_ms,0,blend_radius_m)
  movel([0.524813, -1.268748, -2.641141, -0.802500, 1.570796, 2.095609],accel_mss,speed_ms,0,blend_radius_m)
  movel([0.524669, -1.270323, -2.640263, -0.801803, 1.570796, 2.095466],accel_mss,speed_ms,0,blend_radius_m)
  movel([0.524321, -1.271924, -2.639368, -0.801097, 1.570796, 2.095117],accel_mss,speed_ms,0,blend_radius_m)
  movel([0.523066, -1.275179, -2.637537, -0.799673, 1.570796, 2.093862],accel_mss,speed_ms,0,blend_radius_m)
  movel([0.521175, -1.278426, -2.635698, -0.798265, 1.570796, 2.091972],accel_mss,speed_ms,0,blend_radius_m)
  movel([0.518779, -1.281587, -2.633895, -0.796907, 1.570796, 2.089576],accel_mss,speed_ms,0,blend_radius_m)
  movel([0.516000, -1.284582, -2.632174, -0.795632, 1.570796, 2.086797],accel_mss,speed_ms,0,blend_radius_m)
  movel([0.512959, -1.287337, -2.630582, -0.794470, 1.570796, 2.083755],accel_mss,speed_ms,0,blend_radius_m)
  movel([0.509773, -1.289773, -2.629166, -0.793450, 1.570796, 2.080569],accel_mss,speed_ms,0,blend_radius_m)
  movel([0.506562, -1.291821, -2.627970, -0.792598, 1.570796, 2.077358],accel_mss,speed_ms,0,blend_radius_m)
  movel([0.502578, -1.293812, -2.626802, -0.791775, 1.570796, 2.073374],accel_mss,speed_ms,0,blend_radius_m)
  movel([0.500909, -1.294411, -2.626449, -0.791528, 1.570796, 2.071705],accel_mss,speed_ms,0,blend_radius_m)
  movel([0.499423, -1.294777, -2.626234, -0.791378, 1.570796, 2.070220],accel_mss,speed_ms,0,blend_radius_m)
  movel([0.498100, -1.294930, -2.626144, -0.791315, 1.570796, 2.068896],accel_mss,speed_ms,0,blend_radius_m)
  movel([0.496909, -1.294889, -2.626168, -0.791332, 1.570796, 2.067706],accel_mss,speed_ms,0,blend_radius_m)
  movel([0.494850, -1.294306, -2.626511, -0.791571, 1.570796, 2.065646],accel_mss,speed_ms,0,blend_radius_m)
  movel([0.493058, -1.293197, -2.627163, -0.792029, 1.570796, 2.063855],accel_mss,speed_ms,0,blend_radius_m)
  movel([0.491356, -1.291724, -2.628027, -0.792638, 1.570796, 2.062152],accel_mss,speed_ms,0,blend_radius_m)
  movel([0.487487, -1.288348, -2.629996, -0.794046, 1.570796, 2.058283],accel_mss,speed_ms,0,blend_radius_m)
  movel([0.487259, -1.288202, -2.630080, -0.794107, 1.570796, 2.058055],accel_mss,speed_ms,0,blend_radius_m)
  movel([0.487241, -1.288361, -2.629988, -0.794040, 1.570796, 2.058037],accel_mss,speed_ms,0,blend_radius_m)
  movel([0.487715, -1.289426, -2.629368, -0.793594, 1.570796, 2.058511],accel_mss,speed_ms,0,blend_radius_m)
  movel([0.489967, -1.293431, -2.627026, -0.791932, 1.570796, 2.060763],accel_mss,speed_ms,0,blend_radius_m)
  movel([0.493685, -1.300037, -2.623117, -0.789235, 1.570796, 2.064481],accel_mss,speed_ms,0,blend_radius_m)
  movel([0.489502, -1.298619, -2.623961, -0.789809, 1.570796, 2.060298],accel_mss,speed_ms,0,blend_radius_m)
  movel([0.485053, -1.296746, -2.625072, -0.790572, 1.570796, 2.055849],accel_mss,speed_ms,0,blend_radius_m)
  movel([0.480467, -1.294518, -2.626386, -0.791484, 1.570796, 2.051263],accel_mss,speed_ms,0,blend_radius_m)
  movel([0.475870, -1.292040, -2.627842, -0.792507, 1.570796, 2.046667],accel_mss,speed_ms,0,blend_radius_m)
  movel([0.467201, -1.286704, -2.630949, -0.794736, 1.570796, 2.037997],accel_mss,speed_ms,0,blend_radius_m)
  movel([0.463412, -1.284033, -2.632491, -0.795865, 1.570796, 2.034209],accel_mss,speed_ms,0,blend_radius_m)
  movel([0.460187, -1.281478, -2.633957, -0.796954, 1.570796, 2.030983],accel_mss,speed_ms,0,blend_radius_m)
  movel([0.453118, -1.280912, -2.634280, -0.797196, 1.570796, 2.023914],accel_mss,speed_ms,0,blend_radius_m)
  movel([0.445546, -1.280782, -2.634355, -0.797252, 1.570796, 2.016342],accel_mss,speed_ms,0,blend_radius_m)
  movel([0.429633, -1.281210, -2.634110, -0.797069, 1.570796, 2.000430],accel_mss,speed_ms,0,blend_radius_m)
  movel([0.421650, -1.281457, -2.633969, -0.796963, 1.570796, 1.992447],accel_mss,speed_ms,0,blend_radius_m)
  movel([0.413890, -1.281511, -2.633938, -0.796940, 1.570796, 1.984686],accel_mss,speed_ms,0,blend_radius_m)
  movel([0.406523, -1.281203, -2.634114, -0.797072, 1.570796, 1.977319],accel_mss,speed_ms,0,blend_radius_m)
  movel([0.399719, -1.280368, -2.634591, -0.797429, 1.570796, 1.970515],accel_mss,speed_ms,0,blend_radius_m)
  movel([0.397276, -1.279792, -2.634920, -0.797677, 1.570796, 1.968073],accel_mss,speed_ms,0,blend_radius_m)
  movel([0.395156, -1.279003, -2.635369, -0.798016, 1.570796, 1.965953],accel_mss,speed_ms,0,blend_radius_m)
  movel([0.393364, -1.278012, -2.635933, -0.798444, 1.570796, 1.964160],accel_mss,speed_ms,0,blend_radius_m)
  movel([0.391904, -1.276833, -2.636602, -0.798954, 1.570796, 1.962700],accel_mss,speed_ms,0,blend_radius_m)
  movel([0.390784, -1.275477, -2.637369, -0.799543, 1.570796, 1.961580],accel_mss,speed_ms,0,blend_radius_m)
  movel([0.390006, -1.273960, -2.638224, -0.800205, 1.570796, 1.960802],accel_mss,speed_ms,0,blend_radius_m)
  movel([0.389584, -1.272288, -2.639164, -0.800938, 1.570796, 1.960380],accel_mss,speed_ms,0,blend_radius_m)
  movel([0.389521, -1.270475, -2.640178, -0.801736, 1.570796, 1.960317],accel_mss,speed_ms,0,blend_radius_m)
  movel([0.389824, -1.268539, -2.641257, -0.802593, 1.570796, 1.960621],accel_mss,speed_ms,0,blend_radius_m)
  movel([0.390505, -1.266489, -2.642395, -0.803505, 1.570796, 1.961301],accel_mss,speed_ms,0,blend_radius_m)
  movel([0.391568, -1.264337, -2.643584, -0.804469, 1.570796, 1.962364],accel_mss,speed_ms,0,blend_radius_m)
  movel([0.393021, -1.262102, -2.644812, -0.805475, 1.570796, 1.963817],accel_mss,speed_ms,0,blend_radius_m)
  movel([0.394871, -1.259797, -2.646073, -0.806520, 1.570796, 1.965668],accel_mss,speed_ms,0,blend_radius_m)
  movel([0.397126, -1.257435, -2.647358, -0.807597, 1.570796, 1.967923],accel_mss,speed_ms,0,blend_radius_m)
  movel([0.399795, -1.255035, -2.648656, -0.808698, 1.570796, 1.970591],accel_mss,speed_ms,0,blend_radius_m)
  movel([0.402884, -1.252610, -2.649962, -0.809817, 1.570796, 1.973680],accel_mss,speed_ms,0,blend_radius_m)
  movel([0.402807, -1.255368, -2.648477, -0.808545, 1.570796, 1.973603],accel_mss,speed_ms,0,blend_radius_m)
  movel([0.402862, -1.256664, -2.647776, -0.807949, 1.570796, 1.973658],accel_mss,speed_ms,0,blend_radius_m)
  movel([0.403255, -1.257708, -2.647209, -0.807472, 1.570796, 1.974052],accel_mss,speed_ms,0,blend_radius_m)
  movel([0.403932, -1.258229, -2.646926, -0.807233, 1.570796, 1.974729],accel_mss,speed_ms,0,blend_radius_m)
  movel([0.405026, -1.258589, -2.646731, -0.807069, 1.570796, 1.975822],accel_mss,speed_ms,0,blend_radius_m)
  movel([0.408246, -1.258888, -2.646568, -0.806933, 1.570796, 1.979042],accel_mss,speed_ms,0,blend_radius_m)
  movel([0.412484, -1.258751, -2.646642, -0.806995, 1.570796, 1.983280],accel_mss,speed_ms,0,blend_radius_m)
  movel([0.417321, -1.258316, -2.646879, -0.807194, 1.570796, 1.988117],accel_mss,speed_ms,0,blend_radius_m)
  movel([0.427075, -1.257099, -2.647540, -0.807750, 1.570796, 1.997871],accel_mss,speed_ms,0,blend_radius_m)
  movel([0.434102, -1.256243, -2.648004, -0.808142, 1.570796, 2.004898],accel_mss,speed_ms,0,blend_radius_m)
  movel([0.439885, -1.256053, -2.648106, -0.808230, 1.570796, 2.010681],accel_mss,speed_ms,0,blend_radius_m)
  movel([0.445649, -1.255901, -2.648189, -0.808300, 1.570796, 2.016446],accel_mss,speed_ms,0,blend_radius_m)
  movel([0.439963, -1.249203, -2.651783, -0.811402, 1.570796, 2.010759],accel_mss,speed_ms,0,blend_radius_m)
  movel([0.437249, -1.245447, -2.653776, -0.813166, 1.570796, 2.008045],accel_mss,speed_ms,0,blend_radius_m)
  movel([0.435134, -1.241313, -2.655949, -0.815126, 1.570796, 2.005931],accel_mss,speed_ms,0,blend_radius_m)
  movel([0.434430, -1.239074, -2.657119, -0.816197, 1.570796, 2.005226],accel_mss,speed_ms,0,blend_radius_m)
  movel([0.434026, -1.236701, -2.658350, -0.817337, 1.570796, 2.004822],accel_mss,speed_ms,0,blend_radius_m)
  movel([0.433974, -1.234189, -2.659648, -0.818552, 1.570796, 2.004771],accel_mss,speed_ms,0,blend_radius_m)
  movel([0.434332, -1.231516, -2.661020, -0.819853, 1.570796, 2.005128],accel_mss,speed_ms,0,blend_radius_m)
  movel([0.435146, -1.228674, -2.662470, -0.821245, 1.570796, 2.005942],accel_mss,speed_ms,0,blend_radius_m)
  movel([0.436472, -1.225650, -2.664003, -0.822736, 1.570796, 2.007268],accel_mss,speed_ms,0,blend_radius_m)
  movel([0.438365, -1.222428, -2.665624, -0.824336, 1.570796, 2.009162],accel_mss,speed_ms,0,blend_radius_m)
  movel([0.440881, -1.218999, -2.667337, -0.826053, 1.570796, 2.011678],accel_mss,speed_ms,0,blend_radius_m)
  movel([0.444339, -1.215189, -2.669224, -0.827976, 1.570796, 2.015135],accel_mss,speed_ms,0,blend_radius_m)
  movel([0.448307, -1.211663, -2.670956, -0.829770, 1.570796, 2.019103],accel_mss,speed_ms,0,blend_radius_m)
  movel([0.452636, -1.208516, -2.672490, -0.831383, 1.570796, 2.023432],accel_mss,speed_ms,0,blend_radius_m)
  movel([0.457174, -1.205841, -2.673786, -0.832763, 1.570796, 2.027971],accel_mss,speed_ms,0,blend_radius_m)
  movel([0.461771, -1.203725, -2.674805, -0.833860, 1.570796, 2.032568],accel_mss,speed_ms,0,blend_radius_m)
  movel([0.466271, -1.202267, -2.675503, -0.834618, 1.570796, 2.037067],accel_mss,speed_ms,0,blend_radius_m)
  movel([0.470514, -1.201556, -2.675844, -0.834989, 1.570796, 2.041310],accel_mss,speed_ms,0,blend_radius_m)
  movel([0.474344, -1.201670, -2.675789, -0.834930, 1.570796, 2.045140],accel_mss,speed_ms,0,blend_radius_m)
  movel([0.475997, -1.202348, -2.675465, -0.834576, 1.570796, 2.046793],accel_mss,speed_ms,0,blend_radius_m)
  movel([0.477372, -1.203631, -2.674850, -0.833908, 1.570796, 2.048168],accel_mss,speed_ms,0,blend_radius_m)
  movel([0.477993, -1.205149, -2.674119, -0.833121, 1.570796, 2.048789],accel_mss,speed_ms,0,blend_radius_m)
  movel([0.477872, -1.205884, -2.673765, -0.832740, 1.570796, 2.048669],accel_mss,speed_ms,0,blend_radius_m)
  movel([0.477384, -1.206541, -2.673448, -0.832401, 1.570796, 2.048180],accel_mss,speed_ms,0,blend_radius_m)
  movel([0.476326, -1.205502, -2.673949, -0.832938, 1.570796, 2.047122],accel_mss,speed_ms,0,blend_radius_m)
  movel([0.475227, -1.204827, -2.674274, -0.833288, 1.570796, 2.046024],accel_mss,speed_ms,0,blend_radius_m)
  movel([0.474108, -1.204492, -2.674436, -0.833461, 1.570796, 2.044905],accel_mss,speed_ms,0,blend_radius_m)
  movel([0.472982, -1.204466, -2.674448, -0.833475, 1.570796, 2.043778],accel_mss,speed_ms,0,blend_radius_m)
  movel([0.471863, -1.204725, -2.674323, -0.833340, 1.570796, 2.042659],accel_mss,speed_ms,0,blend_radius_m)
  movel([0.470766, -1.205240, -2.674075, -0.833074, 1.570796, 2.041562],accel_mss,speed_ms,0,blend_radius_m)
  movel([0.469709, -1.205982, -2.673717, -0.832689, 1.570796, 2.040505],accel_mss,speed_ms,0,blend_radius_m)
  movel([0.468709, -1.206920, -2.673264, -0.832205, 1.570796, 2.039506],accel_mss,speed_ms,0,blend_radius_m)
  movel([0.466925, -1.209283, -2.672117, -0.830988, 1.570796, 2.037722],accel_mss,speed_ms,0,blend_radius_m)
  movel([0.465539, -1.212099, -2.670743, -0.829547, 1.570796, 2.036335],accel_mss,speed_ms,0,blend_radius_m)
  movel([0.464652, -1.215154, -2.669241, -0.827993, 1.570796, 2.035448],accel_mss,speed_ms,0,blend_radius_m)
  movel([0.464380, -1.218226, -2.667721, -0.826442, 1.570796, 2.035176],accel_mss,speed_ms,0,blend_radius_m)
  movel([0.464596, -1.219896, -2.666890, -0.825603, 1.570796, 2.035392],accel_mss,speed_ms,0,blend_radius_m)
  movel([0.465144, -1.221725, -2.665977, -0.824687, 1.570796, 2.035940],accel_mss,speed_ms,0,blend_radius_m)
  movel([0.467076, -1.225738, -2.663958, -0.822692, 1.570796, 2.037873],accel_mss,speed_ms,0,blend_radius_m)
  movel([0.469850, -1.230057, -2.661766, -0.820566, 1.570796, 2.040647],accel_mss,speed_ms,0,blend_radius_m)
  movel([0.473145, -1.234459, -2.659509, -0.818421, 1.570796, 2.043941],accel_mss,speed_ms,0,blend_radius_m)
  movel([0.480076, -1.242644, -2.655252, -0.814493, 1.570796, 2.050873],accel_mss,speed_ms,0,blend_radius_m)
  movel([0.485531, -1.248503, -2.652156, -0.811730, 1.570796, 2.056328],accel_mss,speed_ms,0,blend_radius_m)
  movel([0.488288, -1.251408, -2.650606, -0.810375, 1.570796, 2.059085],accel_mss,speed_ms,0,blend_radius_m)
  movel([0.489863, -1.252875, -2.649819, -0.809695, 1.570796, 2.060660],accel_mss,speed_ms,0,blend_radius_m)
  movel([0.491240, -1.253795, -2.649324, -0.809269, 1.570796, 2.062037],accel_mss,speed_ms,0,blend_radius_m)
  movel([0.491732, -1.253917, -2.649259, -0.809213, 1.570796, 2.062529],accel_mss,speed_ms,0,blend_radius_m)
  movel([0.492084, -1.253789, -2.649328, -0.809272, 1.570796, 2.062881],accel_mss,speed_ms,0,blend_radius_m)
  movel([0.492609, -1.252839, -2.649838, -0.809711, 1.570796, 2.063406],accel_mss,speed_ms,0,blend_radius_m)
  movel([0.493352, -1.250069, -2.651322, -0.810998, 1.570796, 2.064148],accel_mss,speed_ms,0,blend_radius_m)
  movel([0.493631, -1.247322, -2.652784, -0.812284, 1.570796, 2.064428],accel_mss,speed_ms,0,blend_radius_m)
  movel([0.493966, -1.241487, -2.655858, -0.815044, 1.570796, 2.064762],accel_mss,speed_ms,0,blend_radius_m)
  movel([0.494616, -1.238193, -2.657576, -0.816619, 1.570796, 2.065413],accel_mss,speed_ms,0,blend_radius_m)
  movel([0.495991, -1.234500, -2.659487, -0.818401, 1.570796, 2.066788],accel_mss,speed_ms,0,blend_radius_m)
  movel([0.497049, -1.232470, -2.660531, -0.819387, 1.570796, 2.067845],accel_mss,speed_ms,0,blend_radius_m)
  movel([0.498407, -1.230297, -2.661643, -0.820449, 1.570796, 2.069203],accel_mss,speed_ms,0,blend_radius_m)
  movel([0.500100, -1.227966, -2.662830, -0.821593, 1.570796, 2.070896],accel_mss,speed_ms,0,blend_radius_m)
  movel([0.502175, -1.225464, -2.664097, -0.822828, 1.570796, 2.072971],accel_mss,speed_ms,0,blend_radius_m)
  movel([0.505211, -1.222364, -2.665657, -0.824369, 1.570796, 2.076007],accel_mss,speed_ms,0,blend_radius_m)
  movel([0.508399, -1.219743, -2.666967, -0.825679, 1.570796, 2.079196],accel_mss,speed_ms,0,blend_radius_m)
  movel([0.511705, -1.217565, -2.668049, -0.826775, 1.570796, 2.082501],accel_mss,speed_ms,0,blend_radius_m)
  movel([0.515093, -1.215790, -2.668928, -0.827671, 1.570796, 2.085889],accel_mss,speed_ms,0,blend_radius_m)
  movel([0.518533, -1.214379, -2.669624, -0.828387, 1.570796, 2.089329],accel_mss,speed_ms,0,blend_radius_m)
  movel([0.521986, -1.213284, -2.670162, -0.828943, 1.570796, 2.092782],accel_mss,speed_ms,0,blend_radius_m)
  movel([0.525425, -1.212463, -2.670564, -0.829361, 1.570796, 2.096221],accel_mss,speed_ms,0,blend_radius_m)
  movel([0.528813, -1.211871, -2.670855, -0.829664, 1.570796, 2.099610],accel_mss,speed_ms,0,blend_radius_m)
  movel([0.534892, -1.211383, -2.671093, -0.829913, 1.570796, 2.105689],accel_mss,speed_ms,0,blend_radius_m)
  movel([0.539796, -1.211691, -2.670942, -0.829755, 1.570796, 2.110593],accel_mss,speed_ms,0,blend_radius_m)
  movel([0.543540, -1.212497, -2.670548, -0.829344, 1.570796, 2.114336],accel_mss,speed_ms,0,blend_radius_m)
  movel([0.546147, -1.213492, -2.670060, -0.828838, 1.570796, 2.116943],accel_mss,speed_ms,0,blend_radius_m)
  movel([0.549455, -1.215604, -2.669019, -0.827765, 1.570796, 2.120252],accel_mss,speed_ms,0,blend_radius_m)
  movel([0.552034, -1.218330, -2.667670, -0.826390, 1.570796, 2.122831],accel_mss,speed_ms,0,blend_radius_m)
  movel([0.553901, -1.221590, -2.666044, -0.824755, 1.570796, 2.124697],accel_mss,speed_ms,0,blend_radius_m)
  movel([0.555071, -1.225305, -2.664177, -0.822907, 1.570796, 2.125867],accel_mss,speed_ms,0,blend_radius_m)
  movel([0.555561, -1.229392, -2.662105, -0.820892, 1.570796, 2.126357],accel_mss,speed_ms,0,blend_radius_m)
  movel([0.555392, -1.233773, -2.659862, -0.818754, 1.570796, 2.126189],accel_mss,speed_ms,0,blend_radius_m)
  movel([0.554582, -1.238380, -2.657479, -0.816530, 1.570796, 2.125378],accel_mss,speed_ms,0,blend_radius_m)
  movel([0.553149, -1.243136, -2.654993, -0.814259, 1.570796, 2.123945],accel_mss,speed_ms,0,blend_radius_m)
  movel([0.551340, -1.247489, -2.652695, -0.812205, 1.570796, 2.122136],accel_mss,speed_ms,0,blend_radius_m)
  movel([0.549252, -1.251811, -2.650390, -0.810188, 1.570796, 2.120048],accel_mss,speed_ms,0,blend_radius_m)
  movel([0.547159, -1.256045, -2.648111, -0.808234, 1.570796, 2.117955],accel_mss,speed_ms,0,blend_radius_m)
  movel([0.545342, -1.260137, -2.645887, -0.806365, 1.570796, 2.116138],accel_mss,speed_ms,0,blend_radius_m)
  movel([0.544073, -1.264026, -2.643755, -0.804608, 1.570796, 2.114869],accel_mss,speed_ms,0,blend_radius_m)
  movel([0.543727, -1.265879, -2.642732, -0.803778, 1.570796, 2.114523],accel_mss,speed_ms,0,blend_radius_m)
  movel([0.543618, -1.267664, -2.641744, -0.802982, 1.570796, 2.114414],accel_mss,speed_ms,0,blend_radius_m)
  movel([0.543780, -1.269371, -2.640794, -0.802224, 1.570796, 2.114577],accel_mss,speed_ms,0,blend_radius_m)
  movel([0.544245, -1.271000, -2.639885, -0.801504, 1.570796, 2.115042],accel_mss,speed_ms,0,blend_radius_m)
  movel([0.545043, -1.272539, -2.639023, -0.800827, 1.570796, 2.115839],accel_mss,speed_ms,0,blend_radius_m)
  movel([0.546209, -1.273988, -2.638208, -0.800193, 1.570796, 2.117005],accel_mss,speed_ms,0,blend_radius_m)
  movel([0.547530, -1.274975, -2.637652, -0.799762, 1.570796, 2.118326],accel_mss,speed_ms,0,blend_radius_m)
  movel([0.549001, -1.275439, -2.637390, -0.799560, 1.570796, 2.119797],accel_mss,speed_ms,0,blend_radius_m)
  movel([0.550573, -1.275448, -2.637385, -0.799556, 1.570796, 2.121370],accel_mss,speed_ms,0,blend_radius_m)
  movel([0.552196, -1.275058, -2.637605, -0.799726, 1.570796, 2.122992],accel_mss,speed_ms,0,blend_radius_m)
  movel([0.553823, -1.274330, -2.638016, -0.800043, 1.570796, 2.124619],accel_mss,speed_ms,0,blend_radius_m)
  movel([0.555400, -1.273326, -2.638580, -0.800482, 1.570796, 2.126196],accel_mss,speed_ms,0,blend_radius_m)
  movel([0.556879, -1.272102, -2.639268, -0.801019, 1.570796, 2.127675],accel_mss,speed_ms,0,blend_radius_m)
  movel([0.558207, -1.270719, -2.640042, -0.801628, 1.570796, 2.129003],accel_mss,speed_ms,0,blend_radius_m)
  movel([0.559334, -1.269239, -2.640868, -0.802282, 1.570796, 2.130130],accel_mss,speed_ms,0,blend_radius_m)
  movel([0.560205, -1.267719, -2.641713, -0.802957, 1.570796, 2.131002],accel_mss,speed_ms,0,blend_radius_m)
  movel([0.560768, -1.266224, -2.642541, -0.803623, 1.570796, 2.131564],accel_mss,speed_ms,0,blend_radius_m)
  movel([0.560969, -1.264812, -2.643322, -0.804255, 1.570796, 2.131765],accel_mss,speed_ms,0,blend_radius_m)
  movel([0.560749, -1.263553, -2.644015, -0.804821, 1.570796, 2.131545],accel_mss,speed_ms,0,blend_radius_m)
  movel([0.560058, -1.262507, -2.644590, -0.805292, 1.570796, 2.130854],accel_mss,speed_ms,0,blend_radius_m)
  movel([0.558841, -1.261738, -2.645011, -0.805639, 1.570796, 2.129638],accel_mss,speed_ms,0,blend_radius_m)
  movel([0.557040, -1.261317, -2.645242, -0.805830, 1.570796, 2.127837],accel_mss,speed_ms,0,blend_radius_m)
  movel([0.557228, -1.262530, -2.644577, -0.805282, 1.570796, 2.128025],accel_mss,speed_ms,0,blend_radius_m)
  movel([0.557104, -1.263706, -2.643931, -0.804752, 1.570796, 2.127900],accel_mss,speed_ms,0,blend_radius_m)
  movel([0.556694, -1.264807, -2.643325, -0.804258, 1.570796, 2.127490],accel_mss,speed_ms,0,blend_radius_m)
  movel([0.556028, -1.265786, -2.642784, -0.803819, 1.570796, 2.126825],accel_mss,speed_ms,0,blend_radius_m)
  movel([0.555130, -1.266614, -2.642326, -0.803449, 1.570796, 2.125926],accel_mss,speed_ms,0,blend_radius_m)
  movel([0.554032, -1.267244, -2.641976, -0.803168, 1.570796, 2.124828],accel_mss,speed_ms,0,blend_radius_m)
  movel([0.552753, -1.267638, -2.641758, -0.802993, 1.570796, 2.123550],accel_mss,speed_ms,0,blend_radius_m)
  movel([0.551323, -1.267762, -2.641689, -0.802938, 1.570796, 2.122119],accel_mss,speed_ms,0,blend_radius_m)
  movel([0.549167, -1.267396, -2.641892, -0.803101, 1.570796, 2.119963],accel_mss,speed_ms,0,blend_radius_m)
  movel([0.547696, -1.266450, -2.642416, -0.803522, 1.570796, 2.118492],accel_mss,speed_ms,0,blend_radius_m)
  movel([0.546860, -1.265004, -2.643216, -0.804169, 1.570796, 2.117656],accel_mss,speed_ms,0,blend_radius_m)
  movel([0.546609, -1.263150, -2.644237, -0.805002, 1.570796, 2.117406],accel_mss,speed_ms,0,blend_radius_m)
  movel([0.546899, -1.260967, -2.645434, -0.805989, 1.570796, 2.117695],accel_mss,speed_ms,0,blend_radius_m)
  movel([0.547678, -1.258546, -2.646754, -0.807089, 1.570796, 2.118475],accel_mss,speed_ms,0,blend_radius_m)
  movel([0.548903, -1.255971, -2.648151, -0.808267, 1.570796, 2.119700],accel_mss,speed_ms,0,blend_radius_m)
  movel([0.550521, -1.253337, -2.649571, -0.809481, 1.570796, 2.121318],accel_mss,speed_ms,0,blend_radius_m)
  movel([0.552491, -1.250731, -2.650968, -0.810690, 1.570796, 2.123287],accel_mss,speed_ms,0,blend_radius_m)
  movel([0.554755, -1.248251, -2.652290, -0.811848, 1.570796, 2.125551],accel_mss,speed_ms,0,blend_radius_m)
  movel([0.557262, -1.245988, -2.653490, -0.812911, 1.570796, 2.128058],accel_mss,speed_ms,0,blend_radius_m)
  movel([0.559958, -1.244045, -2.654515, -0.813828, 1.570796, 2.130755],accel_mss,speed_ms,0,blend_radius_m)
  movel([0.562789, -1.242520, -2.655317, -0.814552, 1.570796, 2.133585],accel_mss,speed_ms,0,blend_radius_m)
  movel([0.565694, -1.241510, -2.655846, -0.815033, 1.570796, 2.136490],accel_mss,speed_ms,0,blend_radius_m)
  movel([0.568617, -1.241113, -2.656054, -0.815222, 1.570796, 2.139414],accel_mss,speed_ms,0,blend_radius_m)
  movel([0.571495, -1.241428, -2.655889, -0.815071, 1.570796, 2.142292],accel_mss,speed_ms,0,blend_radius_m)
  movel([0.573345, -1.242023, -2.655578, -0.814788, 1.570796, 2.144141],accel_mss,speed_ms,0,blend_radius_m)
  movel([0.575004, -1.242834, -2.655152, -0.814403, 1.570796, 2.145801],accel_mss,speed_ms,0,blend_radius_m)
  movel([0.576465, -1.243849, -2.654618, -0.813921, 1.570796, 2.147262],accel_mss,speed_ms,0,blend_radius_m)
  movel([0.577719, -1.245052, -2.653985, -0.813353, 1.570796, 2.148516],accel_mss,speed_ms,0,blend_radius_m)
  movel([0.578762, -1.246430, -2.653256, -0.812703, 1.570796, 2.149558],accel_mss,speed_ms,0,blend_radius_m)
  movel([0.579587, -1.247968, -2.652440, -0.811980, 1.570796, 2.150383],accel_mss,speed_ms,0,blend_radius_m)
  movel([0.580185, -1.249649, -2.651546, -0.811194, 1.570796, 2.150981],accel_mss,speed_ms,0,blend_radius_m)
  movel([0.580553, -1.251461, -2.650578, -0.810350, 1.570796, 2.151350],accel_mss,speed_ms,0,blend_radius_m)
  movel([0.580682, -1.253388, -2.649544, -0.809457, 1.570796, 2.151478],accel_mss,speed_ms,0,blend_radius_m)
  movel([0.580570, -1.255417, -2.648450, -0.808522, 1.570796, 2.151366],accel_mss,speed_ms,0,blend_radius_m)
  movel([0.580210, -1.257533, -2.647304, -0.807551, 1.570796, 2.151006],accel_mss,speed_ms,0,blend_radius_m)
  movel([0.579599, -1.259723, -2.646113, -0.806553, 1.570796, 2.150395],accel_mss,speed_ms,0,blend_radius_m)
  movel([0.578725, -1.261973, -2.644882, -0.805533, 1.570796, 2.149521],accel_mss,speed_ms,0,blend_radius_m)
  movel([0.577588, -1.264270, -2.643621, -0.804499, 1.570796, 2.148384],accel_mss,speed_ms,0,blend_radius_m)
  movel([0.576182, -1.266602, -2.642333, -0.803455, 1.570796, 2.146979],accel_mss,speed_ms,0,blend_radius_m)
  movel([0.574500, -1.268956, -2.641026, -0.802408, 1.570796, 2.145296],accel_mss,speed_ms,0,blend_radius_m)
  movel([0.572448, -1.271109, -2.639824, -0.801456, 1.570796, 2.143244],accel_mss,speed_ms,0,blend_radius_m)
  movel([0.569957, -1.273232, -2.638634, -0.800523, 1.570796, 2.140754],accel_mss,speed_ms,0,blend_radius_m)
  movel([0.567751, -1.274992, -2.637642, -0.799754, 1.570796, 2.138548],accel_mss,speed_ms,0,blend_radius_m)
  movel([0.566551, -1.276060, -2.637039, -0.799290, 1.570796, 2.137348],accel_mss,speed_ms,0,blend_radius_m)
  movel([0.566189, -1.277121, -2.636439, -0.798830, 1.570796, 2.136986],accel_mss,speed_ms,0,blend_radius_m)
  movel([0.565942, -1.278784, -2.635494, -0.798111, 1.570796, 2.136738],accel_mss,speed_ms,0,blend_radius_m)
  movel([0.565676, -1.280612, -2.634452, -0.797325, 1.570796, 2.136473],accel_mss,speed_ms,0,blend_radius_m)
  movel([0.565256, -1.282171, -2.633560, -0.796658, 1.570796, 2.136052],accel_mss,speed_ms,0,blend_radius_m)
  movel([0.564228, -1.284259, -2.632360, -0.795769, 1.570796, 2.135025],accel_mss,speed_ms,0,blend_radius_m)
  movel([0.562995, -1.286188, -2.631247, -0.794954, 1.570796, 2.133791],accel_mss,speed_ms,0,blend_radius_m)
  movel([0.561584, -1.287957, -2.630223, -0.794210, 1.570796, 2.132380],accel_mss,speed_ms,0,blend_radius_m)
  movel([0.560027, -1.289554, -2.629294, -0.793541, 1.570796, 2.130824],accel_mss,speed_ms,0,blend_radius_m)
  movel([0.558350, -1.290977, -2.628464, -0.792948, 1.570796, 2.129146],accel_mss,speed_ms,0,blend_radius_m)
  movel([0.556578, -1.292219, -2.627737, -0.792433, 1.570796, 2.127374],accel_mss,speed_ms,0,blend_radius_m)
  movel([0.554741, -1.293272, -2.627120, -0.791998, 1.570796, 2.125537],accel_mss,speed_ms,0,blend_radius_m)
  movel([0.552865, -1.294134, -2.626613, -0.791642, 1.570796, 2.123662],accel_mss,speed_ms,0,blend_radius_m)
  movel([0.550975, -1.294794, -2.626224, -0.791371, 1.570796, 2.121771],accel_mss,speed_ms,0,blend_radius_m)
  movel([0.549101, -1.295247, -2.625957, -0.791185, 1.570796, 2.119898],accel_mss,speed_ms,0,blend_radius_m)
  movel([0.547267, -1.295484, -2.625817, -0.791088, 1.570796, 2.118063],accel_mss,speed_ms,0,blend_radius_m)
  speed_ms = 0.003
  movel([0.547267, -1.288536, -2.622525, -0.801328, 1.570796, 2.118063],accel_mss,speed_ms,0,blend_radius_m)
  speed_ms = 0.03
  movel([0.547267, -1.261948, -2.609078, -0.841364, 1.570796, 2.118063],accel_mss,speed_ms,0,blend_radius_m)
  #M_RunCode9
  movel([0.552172, -1.270099, -2.604449, -0.837840, 1.570796, 2.122969],accel_mss,speed_ms,0,blend_radius_m)
  #M_RunCode3
  movel([0.552172, -1.296572, -2.617789, -0.798028, 1.570796, 2.122969],accel_mss,speed_ms,0,blend_radius_m)
  speed_ms = 0.003
  movel([0.552172, -1.303485, -2.621054, -0.787849, 1.570796, 2.122969],accel_mss,speed_ms,0,blend_radius_m)
  speed_ms = 0.007
  movel([0.553642, -1.302425, -2.621690, -0.788274, 1.570796, 2.124439],accel_mss,speed_ms,0,blend_radius_m)
  movel([0.556770, -1.300575, -2.622796, -0.789018, 1.570796, 2.127567],accel_mss,speed_ms,0,blend_radius_m)
  movel([0.559771, -1.298669, -2.623931, -0.789789, 1.570796, 2.130567],accel_mss,speed_ms,0,blend_radius_m)
  movel([0.561079, -1.297536, -2.624603, -0.790249, 1.570796, 2.131875],accel_mss,speed_ms,0,blend_radius_m)
  movel([0.562188, -1.296197, -2.625396, -0.790796, 1.570796, 2.132984],accel_mss,speed_ms,0,blend_radius_m)
  movel([0.561646, -1.297257, -2.624769, -0.790363, 1.570796, 2.132442],accel_mss,speed_ms,0,blend_radius_m)
  movel([0.560361, -1.299109, -2.623669, -0.789611, 1.570796, 2.131158],accel_mss,speed_ms,0,blend_radius_m)
  movel([0.558879, -1.300655, -2.622748, -0.788985, 1.570796, 2.129676],accel_mss,speed_ms,0,blend_radius_m)
  movel([0.557252, -1.301999, -2.621945, -0.788445, 1.570796, 2.128048],accel_mss,speed_ms,0,blend_radius_m)
  movel([0.555547, -1.303229, -2.621208, -0.787952, 1.570796, 2.126343],accel_mss,speed_ms,0,blend_radius_m)
  movel([0.552131, -1.305737, -2.619699, -0.786953, 1.570796, 2.122928],accel_mss,speed_ms,0,blend_radius_m)
  movel([0.550547, -1.307202, -2.618814, -0.786374, 1.570796, 2.121343],accel_mss,speed_ms,0,blend_radius_m)
  movel([0.549127, -1.308926, -2.617768, -0.785695, 1.570796, 2.119924],accel_mss,speed_ms,0,blend_radius_m)
  movel([0.547832, -1.310991, -2.616511, -0.784887, 1.570796, 2.118628],accel_mss,speed_ms,0,blend_radius_m)
  movel([0.547226, -1.312110, -2.615827, -0.784452, 1.570796, 2.118023],accel_mss,speed_ms,0,blend_radius_m)
  movel([0.547010, -1.312766, -2.615426, -0.784198, 1.570796, 2.117806],accel_mss,speed_ms,0,blend_radius_m)
  movel([0.547694, -1.313134, -2.615200, -0.784055, 1.570796, 2.118490],accel_mss,speed_ms,0,blend_radius_m)
  movel([0.548220, -1.313474, -2.614991, -0.783924, 1.570796, 2.119017],accel_mss,speed_ms,0,blend_radius_m)
  movel([0.548619, -1.313966, -2.614689, -0.783734, 1.570796, 2.119415],accel_mss,speed_ms,0,blend_radius_m)
  movel([0.549041, -1.315217, -2.613920, -0.783252, 1.570796, 2.119838],accel_mss,speed_ms,0,blend_radius_m)
  movel([0.549102, -1.316317, -2.613241, -0.782830, 1.570796, 2.119899],accel_mss,speed_ms,0,blend_radius_m)
  movel([0.548864, -1.317317, -2.612624, -0.782448, 1.570796, 2.119661],accel_mss,speed_ms,0,blend_radius_m)
  movel([0.548394, -1.318268, -2.612035, -0.782086, 1.570796, 2.119191],accel_mss,speed_ms,0,blend_radius_m)
  movel([0.547005, -1.320232, -2.610815, -0.781342, 1.570796, 2.117802],accel_mss,speed_ms,0,blend_radius_m)
  movel([0.545437, -1.322618, -2.609326, -0.780445, 1.570796, 2.116234],accel_mss,speed_ms,0,blend_radius_m)
  movel([0.543790, -1.325904, -2.607263, -0.779223, 1.570796, 2.114586],accel_mss,speed_ms,0,blend_radius_m)
  movel([0.542270, -1.329169, -2.605198, -0.778022, 1.570796, 2.113066],accel_mss,speed_ms,0,blend_radius_m)
  movel([0.540627, -1.332408, -2.603136, -0.776845, 1.570796, 2.111424],accel_mss,speed_ms,0,blend_radius_m)
  movel([0.538626, -1.335602, -2.601089, -0.775698, 1.570796, 2.109423],accel_mss,speed_ms,0,blend_radius_m)
  movel([0.537326, -1.337268, -2.600015, -0.775105, 1.570796, 2.108122],accel_mss,speed_ms,0,blend_radius_m)
  movel([0.535891, -1.338858, -2.598987, -0.774543, 1.570796, 2.106687],accel_mss,speed_ms,0,blend_radius_m)
  movel([0.532779, -1.341863, -2.597035, -0.773491, 1.570796, 2.103575],accel_mss,speed_ms,0,blend_radius_m)
  movel([0.529582, -1.344732, -2.595160, -0.772497, 1.570796, 2.100378],accel_mss,speed_ms,0,blend_radius_m)
  movel([0.526604, -1.347566, -2.593296, -0.771527, 1.570796, 2.097401],accel_mss,speed_ms,0,blend_radius_m)
  movel([0.522126, -1.352542, -2.589997, -0.769850, 1.570796, 2.092922],accel_mss,speed_ms,0,blend_radius_m)
  movel([0.520258, -1.354690, -2.588562, -0.769136, 1.570796, 2.091054],accel_mss,speed_ms,0,blend_radius_m)
  movel([0.518402, -1.356656, -2.587243, -0.768489, 1.570796, 2.089198],accel_mss,speed_ms,0,blend_radius_m)
  movel([0.516386, -1.358467, -2.586024, -0.767898, 1.570796, 2.087182],accel_mss,speed_ms,0,blend_radius_m)
  movel([0.514033, -1.360159, -2.584880, -0.767349, 1.570796, 2.084829],accel_mss,speed_ms,0,blend_radius_m)
  movel([0.511171, -1.361763, -2.583792, -0.766833, 1.570796, 2.081967],accel_mss,speed_ms,0,blend_radius_m)
  movel([0.507625, -1.363315, -2.582737, -0.766337, 1.570796, 2.078421],accel_mss,speed_ms,0,blend_radius_m)
  movel([0.504731, -1.364316, -2.582054, -0.766019, 1.570796, 2.075528],accel_mss,speed_ms,0,blend_radius_m)
  movel([0.502098, -1.364974, -2.581604, -0.765811, 1.570796, 2.072894],accel_mss,speed_ms,0,blend_radius_m)
  movel([0.499706, -1.365311, -2.581374, -0.765705, 1.570796, 2.070502],accel_mss,speed_ms,0,blend_radius_m)
  movel([0.497545, -1.365349, -2.581348, -0.765693, 1.570796, 2.068342],accel_mss,speed_ms,0,blend_radius_m)
  movel([0.495607, -1.365101, -2.581517, -0.765771, 1.570796, 2.066404],accel_mss,speed_ms,0,blend_radius_m)
  movel([0.493880, -1.364592, -2.581865, -0.765932, 1.570796, 2.064677],accel_mss,speed_ms,0,blend_radius_m)
  movel([0.492350, -1.363836, -2.582381, -0.766171, 1.570796, 2.063146],accel_mss,speed_ms,0,blend_radius_m)
  movel([0.491008, -1.362853, -2.583051, -0.766485, 1.570796, 2.061804],accel_mss,speed_ms,0,blend_radius_m)
  movel([0.489847, -1.361664, -2.583860, -0.766865, 1.570796, 2.060643],accel_mss,speed_ms,0,blend_radius_m)
  movel([0.488853, -1.360286, -2.584795, -0.767309, 1.570796, 2.059649],accel_mss,speed_ms,0,blend_radius_m)
  movel([0.487336, -1.357033, -2.586990, -0.768366, 1.570796, 2.058132],accel_mss,speed_ms,0,blend_radius_m)
  movel([0.486384, -1.353244, -2.589529, -0.769616, 1.570796, 2.057180],accel_mss,speed_ms,0,blend_radius_m)
  movel([0.485926, -1.349068, -2.592304, -0.771017, 1.570796, 2.056722],accel_mss,speed_ms,0,blend_radius_m)
  movel([0.485948, -1.344902, -2.595048, -0.772438, 1.570796, 2.056744],accel_mss,speed_ms,0,blend_radius_m)
  movel([0.486105, -1.339479, -2.598585, -0.774325, 1.570796, 2.056901],accel_mss,speed_ms,0,blend_radius_m)
  movel([0.485987, -1.333551, -2.602405, -0.776433, 1.570796, 2.056783],accel_mss,speed_ms,0,blend_radius_m)
  movel([0.485696, -1.330637, -2.604265, -0.777487, 1.570796, 2.056492],accel_mss,speed_ms,0,blend_radius_m)
  movel([0.485177, -1.327893, -2.606007, -0.778489, 1.570796, 2.055973],accel_mss,speed_ms,0,blend_radius_m)
  movel([0.484377, -1.325421, -2.607567, -0.779401, 1.570796, 2.055173],accel_mss,speed_ms,0,blend_radius_m)
  movel([0.483243, -1.323321, -2.608885, -0.780182, 1.570796, 2.054039],accel_mss,speed_ms,0,blend_radius_m)
  movel([0.481721, -1.321700, -2.609899, -0.780789, 1.570796, 2.052517],accel_mss,speed_ms,0,blend_radius_m)
  movel([0.479761, -1.320661, -2.610548, -0.781180, 1.570796, 2.050557],accel_mss,speed_ms,0,blend_radius_m)
  movel([0.478597, -1.320395, -2.610713, -0.781281, 1.570796, 2.049394],accel_mss,speed_ms,0,blend_radius_m)
  movel([0.477308, -1.320313, -2.610765, -0.781312, 1.570796, 2.048104],accel_mss,speed_ms,0,blend_radius_m)
  movel([0.475881, -1.320429, -2.610692, -0.781268, 1.570796, 2.046678],accel_mss,speed_ms,0,blend_radius_m)
  movel([0.474318, -1.320753, -2.610490, -0.781146, 1.570796, 2.045115],accel_mss,speed_ms,0,blend_radius_m)
  movel([0.472608, -1.321301, -2.610148, -0.780939, 1.570796, 2.043404],accel_mss,speed_ms,0,blend_radius_m)
  movel([0.470748, -1.322082, -2.609661, -0.780646, 1.570796, 2.041545],accel_mss,speed_ms,0,blend_radius_m)
  movel([0.466556, -1.324398, -2.608210, -0.779781, 1.570796, 2.037353],accel_mss,speed_ms,0,blend_radius_m)
  movel([0.464696, -1.325888, -2.607273, -0.779228, 1.570796, 2.035492],accel_mss,speed_ms,0,blend_radius_m)
  movel([0.462981, -1.327628, -2.606174, -0.778587, 1.570796, 2.033777],accel_mss,speed_ms,0,blend_radius_m)
  movel([0.461442, -1.329614, -2.604916, -0.777859, 1.570796, 2.032238],accel_mss,speed_ms,0,blend_radius_m)
  movel([0.460112, -1.331836, -2.603502, -0.777052, 1.570796, 2.030908],accel_mss,speed_ms,0,blend_radius_m)
  movel([0.462912, -1.330818, -2.604150, -0.777421, 1.570796, 2.033708],accel_mss,speed_ms,0,blend_radius_m)
  movel([0.465588, -1.330111, -2.604600, -0.777678, 1.570796, 2.036384],accel_mss,speed_ms,0,blend_radius_m)
  movel([0.468124, -1.329702, -2.604860, -0.777827, 1.570796, 2.038920],accel_mss,speed_ms,0,blend_radius_m)
  movel([0.470505, -1.329588, -2.604932, -0.777869, 1.570796, 2.041302],accel_mss,speed_ms,0,blend_radius_m)
  movel([0.472715, -1.329757, -2.604825, -0.777807, 1.570796, 2.043511],accel_mss,speed_ms,0,blend_radius_m)
  movel([0.474741, -1.330196, -2.604546, -0.777647, 1.570796, 2.045537],accel_mss,speed_ms,0,blend_radius_m)
  movel([0.476564, -1.330900, -2.604098, -0.777391, 1.570796, 2.047360],accel_mss,speed_ms,0,blend_radius_m)
  movel([0.478174, -1.331852, -2.603491, -0.777046, 1.570796, 2.048970],accel_mss,speed_ms,0,blend_radius_m)
  movel([0.479552, -1.333048, -2.602727, -0.776614, 1.570796, 2.050348],accel_mss,speed_ms,0,blend_radius_m)
  movel([0.480692, -1.334469, -2.601817, -0.776103, 1.570796, 2.051488],accel_mss,speed_ms,0,blend_radius_m)
  movel([0.481577, -1.336106, -2.600765, -0.775519, 1.570796, 2.052373],accel_mss,speed_ms,0,blend_radius_m)
  movel([0.482196, -1.337947, -2.599577, -0.774865, 1.570796, 2.052992],accel_mss,speed_ms,0,blend_radius_m)
  movel([0.482536, -1.339978, -2.598261, -0.774149, 1.570796, 2.053332],accel_mss,speed_ms,0,blend_radius_m)
  movel([0.482587, -1.342191, -2.596822, -0.773377, 1.570796, 2.053383],accel_mss,speed_ms,0,blend_radius_m)
  movel([0.482337, -1.344570, -2.595266, -0.772553, 1.570796, 2.053133],accel_mss,speed_ms,0,blend_radius_m)
  movel([0.481778, -1.347105, -2.593600, -0.771684, 1.570796, 2.052575],accel_mss,speed_ms,0,blend_radius_m)
  movel([0.481091, -1.349237, -2.592192, -0.770960, 1.570796, 2.051888],accel_mss,speed_ms,0,blend_radius_m)
  movel([0.480231, -1.351313, -2.590815, -0.770261, 1.570796, 2.051027],accel_mss,speed_ms,0,blend_radius_m)
  movel([0.479210, -1.353326, -2.589474, -0.769589, 1.570796, 2.050006],accel_mss,speed_ms,0,blend_radius_m)
  movel([0.478047, -1.355269, -2.588175, -0.768945, 1.570796, 2.048843],accel_mss,speed_ms,0,blend_radius_m)
  movel([0.475338, -1.358930, -2.585712, -0.767748, 1.570796, 2.046134],accel_mss,speed_ms,0,blend_radius_m)
  movel([0.472212, -1.362252, -2.583460, -0.766677, 1.570796, 2.043009],accel_mss,speed_ms,0,blend_radius_m)
  movel([0.468777, -1.365196, -2.581452, -0.765741, 1.570796, 2.039574],accel_mss,speed_ms,0,blend_radius_m)
  movel([0.465138, -1.367719, -2.579722, -0.764949, 1.570796, 2.035934],accel_mss,speed_ms,0,blend_radius_m)
  movel([0.461390, -1.369783, -2.578299, -0.764307, 1.570796, 2.032186],accel_mss,speed_ms,0,blend_radius_m)
  movel([0.457636, -1.371342, -2.577221, -0.763826, 1.570796, 2.028432],accel_mss,speed_ms,0,blend_radius_m)
  movel([0.453973, -1.372354, -2.576519, -0.763516, 1.570796, 2.024770],accel_mss,speed_ms,0,blend_radius_m)
  movel([0.450502, -1.372775, -2.576227, -0.763388, 1.570796, 2.021298],accel_mss,speed_ms,0,blend_radius_m)
  movel([0.447318, -1.372554, -2.576380, -0.763455, 1.570796, 2.018114],accel_mss,speed_ms,0,blend_radius_m)
  movel([0.445864, -1.372189, -2.576633, -0.763567, 1.570796, 2.016660],accel_mss,speed_ms,0,blend_radius_m)
  movel([0.444520, -1.371643, -2.577012, -0.763734, 1.570796, 2.015316],accel_mss,speed_ms,0,blend_radius_m)
  movel([0.443297, -1.370913, -2.577518, -0.763958, 1.570796, 2.014093],accel_mss,speed_ms,0,blend_radius_m)
  movel([0.442210, -1.369986, -2.578159, -0.764244, 1.570796, 2.013006],accel_mss,speed_ms,0,blend_radius_m)
  movel([0.441269, -1.368858, -2.578937, -0.764594, 1.570796, 2.012065],accel_mss,speed_ms,0,blend_radius_m)
  movel([0.440490, -1.367522, -2.579857, -0.765010, 1.570796, 2.011286],accel_mss,speed_ms,0,blend_radius_m)
  movel([0.439886, -1.365971, -2.580922, -0.765496, 1.570796, 2.010682],accel_mss,speed_ms,0,blend_radius_m)
  movel([0.439471, -1.364192, -2.582138, -0.766058, 1.570796, 2.010267],accel_mss,speed_ms,0,blend_radius_m)
  movel([0.439257, -1.362180, -2.583509, -0.766700, 1.570796, 2.010053],accel_mss,speed_ms,0,blend_radius_m)
  movel([0.439261, -1.359925, -2.585039, -0.767425, 1.570796, 2.010057],accel_mss,speed_ms,0,blend_radius_m)
  movel([0.439580, -1.357972, -2.586358, -0.768059, 1.570796, 2.010377],accel_mss,speed_ms,0,blend_radius_m)
  movel([0.440970, -1.352415, -2.590082, -0.769892, 1.570796, 2.011766],accel_mss,speed_ms,0,blend_radius_m)
  movel([0.442275, -1.348414, -2.592736, -0.771238, 1.570796, 2.013072],accel_mss,speed_ms,0,blend_radius_m)
  movel([0.444102, -1.343666, -2.595858, -0.772865, 1.570796, 2.014898],accel_mss,speed_ms,0,blend_radius_m)
  movel([0.446548, -1.338213, -2.599405, -0.774771, 1.570796, 2.017345],accel_mss,speed_ms,0,blend_radius_m)
  movel([0.449703, -1.332104, -2.603330, -0.776955, 1.570796, 2.020499],accel_mss,speed_ms,0,blend_radius_m)
  movel([0.452244, -1.327821, -2.606052, -0.778516, 1.570796, 2.023040],accel_mss,speed_ms,0,blend_radius_m)
  movel([0.454869, -1.323977, -2.608474, -0.779938, 1.570796, 2.025665],accel_mss,speed_ms,0,blend_radius_m)
  movel([0.457540, -1.320552, -2.610616, -0.781221, 1.570796, 2.028337],accel_mss,speed_ms,0,blend_radius_m)
  movel([0.460225, -1.317531, -2.612491, -0.782367, 1.570796, 2.031021],accel_mss,speed_ms,0,blend_radius_m)
  movel([0.462887, -1.314896, -2.614118, -0.783376, 1.570796, 2.033683],accel_mss,speed_ms,0,blend_radius_m)
  movel([0.465492, -1.312622, -2.615514, -0.784254, 1.570796, 2.036288],accel_mss,speed_ms,0,blend_radius_m)
  movel([0.468006, -1.310685, -2.616697, -0.785007, 1.570796, 2.038803],accel_mss,speed_ms,0,blend_radius_m)
  movel([0.470395, -1.309067, -2.617682, -0.785640, 1.570796, 2.041191],accel_mss,speed_ms,0,blend_radius_m)
  movel([0.474657, -1.306676, -2.619132, -0.786582, 1.570796, 2.045454],accel_mss,speed_ms,0,blend_radius_m)
  movel([0.478017, -1.305243, -2.619997, -0.787149, 1.570796, 2.048813],accel_mss,speed_ms,0,blend_radius_m)
  movel([0.480213, -1.304549, -2.620415, -0.787425, 1.570796, 2.051009],accel_mss,speed_ms,0,blend_radius_m)
  movel([0.481000, -1.304368, -2.620524, -0.787498, 1.570796, 2.051796],accel_mss,speed_ms,0,blend_radius_m)
  movel([0.484601, -1.303814, -2.620857, -0.787718, 1.570796, 2.055397],accel_mss,speed_ms,0,blend_radius_m)
